FUNCTION_BLOCK "RD_PR_GantryUnload_Seqv25"   // FB2, LAD
VERSION : 0.1
// stored: AutoNumber true, IsIECCheckEnabled false, UDAEnableTagReadback false
   VAR_INPUT
      iAutoRunning : Bool;
      iCenteringSlideAtHome : Bool;
      iCenteringSlideAtWork : Bool;
      iDistSenHighLimit : Int;
      iDistSenLowLimit : Int;
      iDistSensorIP : Int;
      iDryCycleWithoutPal : Bool;
      iGantryOutofZone : Bool;
      iGantryPickOver : Bool;
      iPCAckZero : Bool;
      iPCBypass : Bool;
      iPCDataReadOver : Bool;
      iPCDataWriteOver : Bool;
      iPalletPresent : Bool;
      iProcessStart : Bool;
      iReset_fault : Bool;
      iRetryPB : Bool;
      iScanErr : Bool;
      iScanOver : Bool;
      iScannerBypass : Bool;
      iSstMode : Bool;
      iSstPB : Bool;
   END_VAR
   VAR_OUTPUT
      qCenteringSlideAdvance : Bool;
      qCenteringSlideRetract : Bool;
      qCheckDistance : Bool;
      qGantryOkToUnload : Bool;
      qMsg : Array[0..2] of Bool;
      qPCReadCmd : Bool;
      qPCUploadCmd : Bool;
      qProcessOver : Bool;
      qScanCmd : Bool;
   END_VAR
   VAR DB_SPECIFIC
      StateNo : Int;
      s44_WaitResetRelease : Bool;
      s44_WaitResetRelease_T1 : Bool;
      s45_WaitGantryOutZone : Bool;
      s45_WaitGantryOutZone_T1 : Bool;
      s46_ChkStationHome : Bool;
      s46_ChkStationHome_T1 : Bool;
      s46_ChkStationHome_T2 : Bool;
      s47_WaitProcStartPZR : Bool;
      s47_WaitProcStartPZR_T1 : Bool;
      s48_ChkRecovery : Bool;
      s48_ChkRecovery_T1 : Bool;
      s48_ChkRecovery_T2 : Bool;
      s48_ChkRecovery_T3 : Bool;
      s49_WaitCentSlideAdv : Bool;
      s49_WaitCentSlideAdv_T1 : Bool;
      s50_WaitDistSensorFB : Bool;
      s50_WaitDistSensorFB_T1 : Bool;
      s51_WaitCentSlideRet : Bool;
      s51_WaitCentSlideRet_T1 : Bool;
      s52_WaitScanOver : Bool;
      s52_WaitScanOver_T1 : Bool;
      s52_WaitScanOver_T2 : Bool;
      s53_ChkDistOkWithPC : Bool;
      s53_ChkDistOkWithPC_T1 : Bool;
      s53_ChkDistOkWithPC_T2 : Bool;
      s54_WaitGantryUnload : Bool;
      s54_WaitGantryUnload_T1 : Bool;
      s55_WaitGantryUnldOvr : Bool;
      s55_WaitGantryUnldOvr_T1 : Bool;
      s56_WaitGantryOutZone : Bool;
      s56_WaitGantryOutZone_T1 : Bool;
      s57_ChkReelAbsentConv : Bool;
      s57_ChkReelAbsentConv_T1 : Bool;
      s58_WaitProcStartLow : Bool;
      s58_WaitProcStartLow_T1 : Bool;
      s61_ChkMeasDiamTol : Bool;
      s61_ChkMeasDiamTol_T1 : Bool;
      s61_ChkMeasDiamTol_T2 : Bool;
      s62_WaitPCAckZero : Bool;
      s62_WaitPCAckZero_T1 : Bool;
      s63_WaitDataWritePC : Bool;
      s63_WaitDataWritePC_T1 : Bool;
      s64_WaitOperatorIntv : Bool;
      s64_WaitOperatorIntv_T1 : Bool;
      s65_ChkScanRetryOver : Bool;
      s65_ChkScanRetryOver_T1 : Bool;
      s65_ChkScanRetryOver_T2 : Bool;
      s66_WaitOperatorDecis : Bool;
      s66_WaitOperatorDecis_T1 : Bool;
      s67_WaitCentSlideRet : Bool;
      s67_WaitCentSlideRet_T1 : Bool;
      s68_WaitPCAckZeroRead : Bool;
      s68_WaitPCAckZeroRead_T1 : Bool;
      s69_WaitDataReadPC : Bool;
      s69_WaitDataReadPC_T1 : Bool;
      sDistanceHighLimit : Int;
      sDistanceLowLimit : Int;
      sRecoveryInt : Int;
      sScanRetryCount : Int;
      sSst : Bool;
      sSstPulse : Bool;
      sSstRise : Bool;
   END_VAR
   VAR_TEMP
      tOne : Bool;
   END_VAR
   VAR_TEMP   // added for the SCL form of the ladder/FBD networks
      _w1 : Bool;
   END_VAR
BEGIN

REGION Network 1
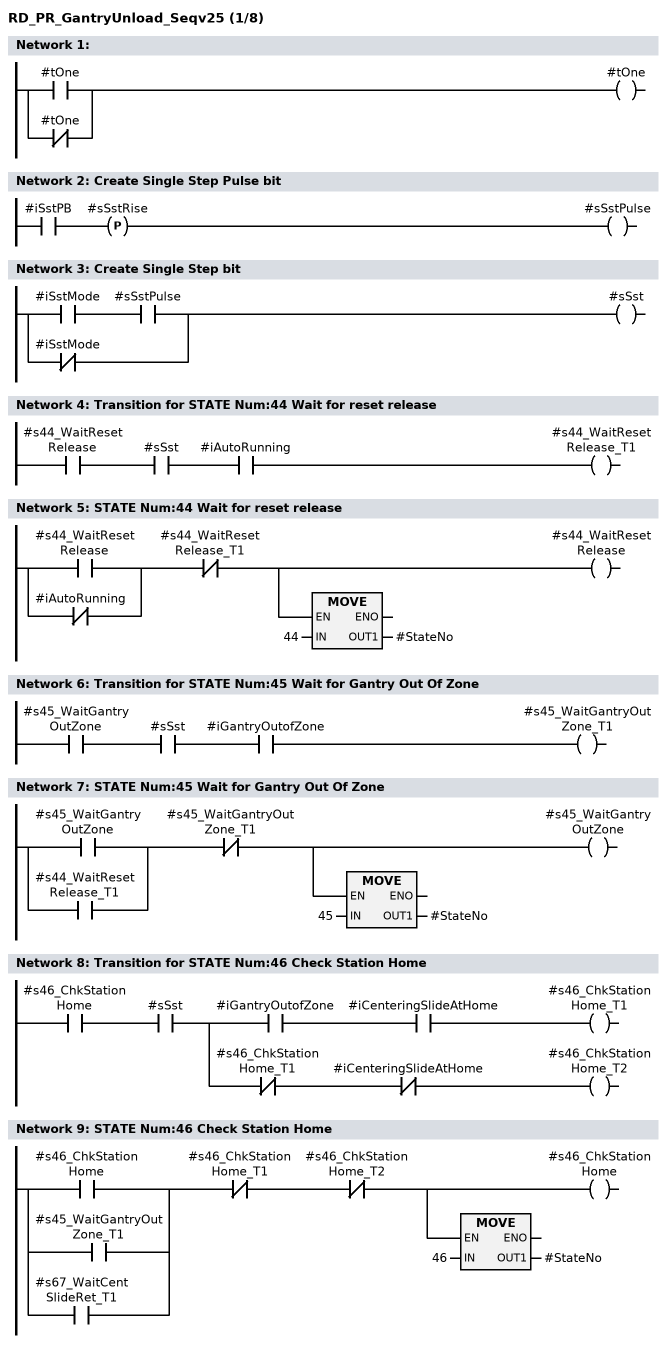
   RUNG wire#powerrail
      Contact( #tOne )
      wire#w1
      Coil( #tOne )
   END_RUNG
   RUNG wire#powerrail
      I_Contact( #tOne )
   END_RUNG wire#w1
   // the same network as SCL:
   #tOne := #tOne OR NOT #tOne;
END_REGION

REGION Network 2: Create Single Step Pulse bit
   RUNG wire#powerrail
      Contact( #iSstPB )
      P_Trig( #sSstRise )
      Coil( #sSstPulse )
   END_RUNG
   // the same network as SCL:
   #_w1 := #iSstPB AND NOT #sSstRise;   // rising edge
   #sSstRise := #iSstPB;
   #sSstPulse := #_w1;
END_REGION

REGION Network 3: Create Single Step bit
   RUNG wire#powerrail
      Contact( #iSstMode )
      Contact( #sSstPulse )
      wire#w1
      Coil( #sSst )
   END_RUNG
   RUNG wire#powerrail
      I_Contact( #iSstMode )
   END_RUNG wire#w1
   // the same network as SCL:
   #sSst := (#iSstMode AND #sSstPulse) OR NOT #iSstMode;
END_REGION

REGION Network 4: Transition for STATE Num:44 Wait for reset release
   RUNG wire#powerrail
      Contact( #s44_WaitResetRelease )
      Contact( #sSst )
      Contact( #iAutoRunning )
      Coil( #s44_WaitResetRelease_T1 )
   END_RUNG
   // the same network as SCL:
   #s44_WaitResetRelease_T1 := #s44_WaitResetRelease AND #sSst AND #iAutoRunning;
END_REGION

REGION Network 5: STATE Num:44 Wait for reset release
   RUNG wire#powerrail
      Contact( #s44_WaitResetRelease )
      wire#w1
      I_Contact( #s44_WaitResetRelease_T1 )
      wire#w2
      Coil( #s44_WaitResetRelease )
   END_RUNG
   RUNG wire#powerrail
      I_Contact( #iAutoRunning )
   END_RUNG wire#w1
   RUNG wire#w2
      { S7_GenerateENO := "TRUE" } Move(in := 44, out1 => #StateNo)
   END_RUNG
   // the same network as SCL:
   #s44_WaitResetRelease := (#s44_WaitResetRelease OR NOT #iAutoRunning) AND NOT #s44_WaitResetRelease_T1;
   IF #s44_WaitResetRelease THEN #StateNo := 44; END_IF;
END_REGION

REGION Network 6: Transition for STATE Num:45 Wait for Gantry Out Of Zone
   RUNG wire#powerrail
      Contact( #s45_WaitGantryOutZone )
      Contact( #sSst )
      Contact( #iGantryOutofZone )
      Coil( #s45_WaitGantryOutZone_T1 )
   END_RUNG
   // the same network as SCL:
   #s45_WaitGantryOutZone_T1 := #s45_WaitGantryOutZone AND #sSst AND #iGantryOutofZone;
END_REGION

REGION Network 7: STATE Num:45 Wait for Gantry Out Of Zone
   RUNG wire#powerrail
      Contact( #s45_WaitGantryOutZone )
      wire#w1
      I_Contact( #s45_WaitGantryOutZone_T1 )
      wire#w2
      Coil( #s45_WaitGantryOutZone )
   END_RUNG
   RUNG wire#powerrail
      Contact( #s44_WaitResetRelease_T1 )
   END_RUNG wire#w1
   RUNG wire#w2
      { S7_GenerateENO := "TRUE" } Move(in := 45, out1 => #StateNo)
   END_RUNG
   // the same network as SCL:
   #s45_WaitGantryOutZone := (#s45_WaitGantryOutZone OR #s44_WaitResetRelease_T1) AND NOT #s45_WaitGantryOutZone_T1;
   IF #s45_WaitGantryOutZone THEN #StateNo := 45; END_IF;
END_REGION

REGION Network 8: Transition for STATE Num:46 Check Station Home
   RUNG wire#powerrail
      Contact( #s46_ChkStationHome )
      Contact( #sSst )
      wire#w1
      Contact( #iGantryOutofZone )
      Contact( #iCenteringSlideAtHome )
      Coil( #s46_ChkStationHome_T1 )
   END_RUNG
   RUNG wire#w1
      I_Contact( #s46_ChkStationHome_T1 )
      I_Contact( #iCenteringSlideAtHome )
      Coil( #s46_ChkStationHome_T2 )
   END_RUNG
   // the same network as SCL:
   #_w1 := #s46_ChkStationHome AND #sSst;
   #s46_ChkStationHome_T1 := #_w1 AND #iGantryOutofZone AND #iCenteringSlideAtHome;
   #s46_ChkStationHome_T2 := #_w1 AND NOT #s46_ChkStationHome_T1 AND NOT #iCenteringSlideAtHome;
END_REGION

REGION Network 9: STATE Num:46 Check Station Home
   RUNG wire#powerrail
      Contact( #s46_ChkStationHome )
      wire#w1
      I_Contact( #s46_ChkStationHome_T1 )
      I_Contact( #s46_ChkStationHome_T2 )
      wire#w2
      Coil( #s46_ChkStationHome )
   END_RUNG
   RUNG wire#powerrail
      Contact( #s45_WaitGantryOutZone_T1 )
   END_RUNG wire#w1
   RUNG wire#powerrail
      Contact( #s67_WaitCentSlideRet_T1 )
   END_RUNG wire#w1
   RUNG wire#w2
      { S7_GenerateENO := "TRUE" } Move(in := 46, out1 => #StateNo)
   END_RUNG
   // the same network as SCL:
   #s46_ChkStationHome := (#s46_ChkStationHome OR #s45_WaitGantryOutZone_T1 OR #s67_WaitCentSlideRet_T1) AND NOT #s46_ChkStationHome_T1 AND NOT #s46_ChkStationHome_T2;
   IF #s46_ChkStationHome THEN #StateNo := 46; END_IF;
END_REGION

REGION Network 10: Transition for STATE Num:47 Wait for Process Start From PZR
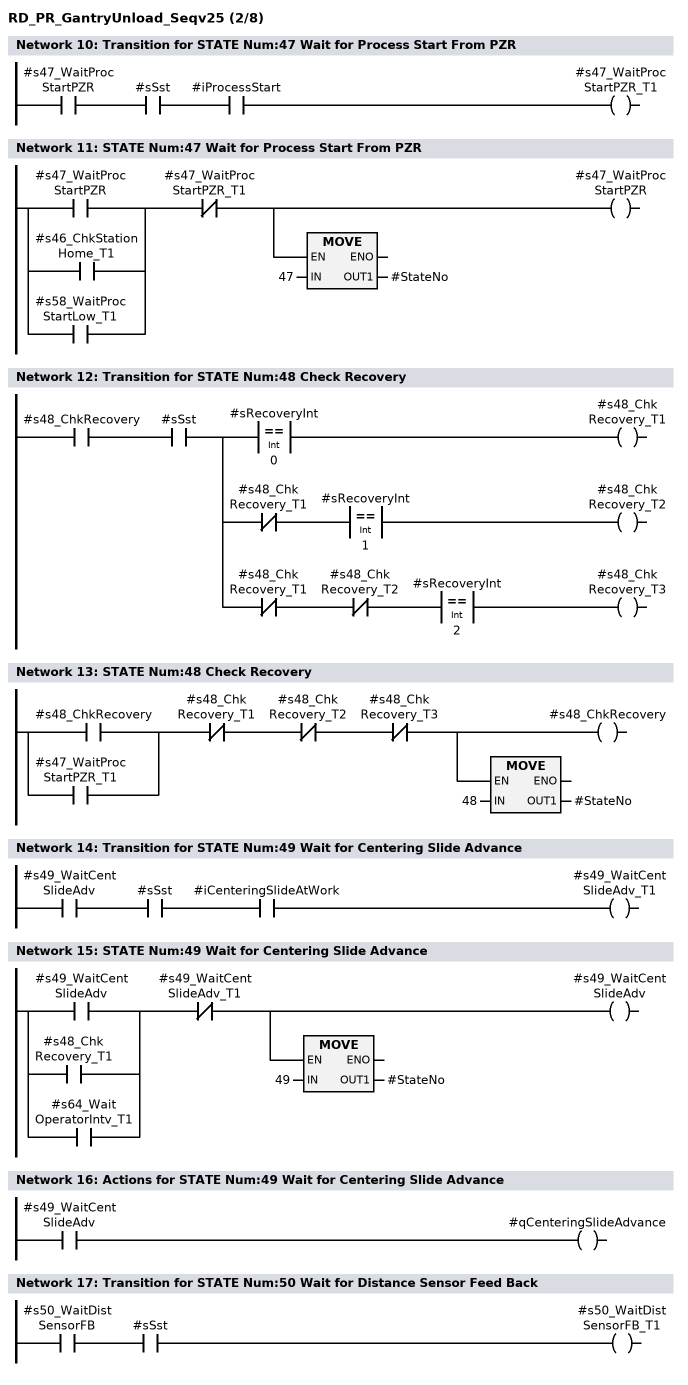
   RUNG wire#powerrail
      Contact( #s47_WaitProcStartPZR )
      Contact( #sSst )
      Contact( #iProcessStart )
      Coil( #s47_WaitProcStartPZR_T1 )
   END_RUNG
   // the same network as SCL:
   #s47_WaitProcStartPZR_T1 := #s47_WaitProcStartPZR AND #sSst AND #iProcessStart;
END_REGION

REGION Network 11: STATE Num:47 Wait for Process Start From PZR
   RUNG wire#powerrail
      Contact( #s47_WaitProcStartPZR )
      wire#w1
      I_Contact( #s47_WaitProcStartPZR_T1 )
      wire#w2
      Coil( #s47_WaitProcStartPZR )
   END_RUNG
   RUNG wire#powerrail
      Contact( #s46_ChkStationHome_T1 )
   END_RUNG wire#w1
   RUNG wire#powerrail
      Contact( #s58_WaitProcStartLow_T1 )
   END_RUNG wire#w1
   RUNG wire#w2
      { S7_GenerateENO := "TRUE" } Move(in := 47, out1 => #StateNo)
   END_RUNG
   // the same network as SCL:
   #s47_WaitProcStartPZR := (#s47_WaitProcStartPZR OR #s46_ChkStationHome_T1 OR #s58_WaitProcStartLow_T1) AND NOT #s47_WaitProcStartPZR_T1;
   IF #s47_WaitProcStartPZR THEN #StateNo := 47; END_IF;
END_REGION

REGION Network 12: Transition for STATE Num:48 Check Recovery
   RUNG wire#powerrail
      Contact( #s48_ChkRecovery )
      Contact( #sSst )
      wire#w1
      { S7_Templates := "SrcType := Int" } EQ_Contact(in1 := #sRecoveryInt, in2 := 0)
      Coil( #s48_ChkRecovery_T1 )
   END_RUNG
   RUNG wire#w1
      I_Contact( #s48_ChkRecovery_T1 )
      { S7_Templates := "SrcType := Int" } EQ_Contact(in1 := #sRecoveryInt, in2 := 1)
      Coil( #s48_ChkRecovery_T2 )
   END_RUNG
   RUNG wire#w1
      I_Contact( #s48_ChkRecovery_T1 )
      I_Contact( #s48_ChkRecovery_T2 )
      { S7_Templates := "SrcType := Int" } EQ_Contact(in1 := #sRecoveryInt, in2 := 2)
      Coil( #s48_ChkRecovery_T3 )
   END_RUNG
   // the same network as SCL:
   #_w1 := #s48_ChkRecovery AND #sSst;
   #s48_ChkRecovery_T1 := #_w1 AND (#sRecoveryInt = 0);
   #s48_ChkRecovery_T2 := #_w1 AND NOT #s48_ChkRecovery_T1 AND (#sRecoveryInt = 1);
   #s48_ChkRecovery_T3 := #_w1 AND NOT #s48_ChkRecovery_T1 AND NOT #s48_ChkRecovery_T2 AND (#sRecoveryInt = 2);
END_REGION

REGION Network 13: STATE Num:48 Check Recovery
   RUNG wire#powerrail
      Contact( #s48_ChkRecovery )
      wire#w1
      I_Contact( #s48_ChkRecovery_T1 )
      I_Contact( #s48_ChkRecovery_T2 )
      I_Contact( #s48_ChkRecovery_T3 )
      wire#w2
      Coil( #s48_ChkRecovery )
   END_RUNG
   RUNG wire#powerrail
      Contact( #s47_WaitProcStartPZR_T1 )
   END_RUNG wire#w1
   RUNG wire#w2
      { S7_GenerateENO := "TRUE" } Move(in := 48, out1 => #StateNo)
   END_RUNG
   // the same network as SCL:
   #s48_ChkRecovery := (#s48_ChkRecovery OR #s47_WaitProcStartPZR_T1) AND NOT #s48_ChkRecovery_T1 AND NOT #s48_ChkRecovery_T2 AND NOT #s48_ChkRecovery_T3;
   IF #s48_ChkRecovery THEN #StateNo := 48; END_IF;
END_REGION

REGION Network 14: Transition for STATE Num:49 Wait for Centering Slide Advance
   RUNG wire#powerrail
      Contact( #s49_WaitCentSlideAdv )
      Contact( #sSst )
      Contact( #iCenteringSlideAtWork )
      Coil( #s49_WaitCentSlideAdv_T1 )
   END_RUNG
   // the same network as SCL:
   #s49_WaitCentSlideAdv_T1 := #s49_WaitCentSlideAdv AND #sSst AND #iCenteringSlideAtWork;
END_REGION

REGION Network 15: STATE Num:49 Wait for Centering Slide Advance
   RUNG wire#powerrail
      Contact( #s49_WaitCentSlideAdv )
      wire#w1
      I_Contact( #s49_WaitCentSlideAdv_T1 )
      wire#w2
      Coil( #s49_WaitCentSlideAdv )
   END_RUNG
   RUNG wire#powerrail
      Contact( #s48_ChkRecovery_T1 )
   END_RUNG wire#w1
   RUNG wire#powerrail
      Contact( #s64_WaitOperatorIntv_T1 )
   END_RUNG wire#w1
   RUNG wire#w2
      { S7_GenerateENO := "TRUE" } Move(in := 49, out1 => #StateNo)
   END_RUNG
   // the same network as SCL:
   #s49_WaitCentSlideAdv := (#s49_WaitCentSlideAdv OR #s48_ChkRecovery_T1 OR #s64_WaitOperatorIntv_T1) AND NOT #s49_WaitCentSlideAdv_T1;
   IF #s49_WaitCentSlideAdv THEN #StateNo := 49; END_IF;
END_REGION

REGION Network 16: Actions for STATE Num:49 Wait for Centering Slide Advance
   RUNG wire#powerrail
      Contact( #s49_WaitCentSlideAdv )
      Coil( #qCenteringSlideAdvance )
   END_RUNG
   // the same network as SCL:
   #qCenteringSlideAdvance := #s49_WaitCentSlideAdv;
END_REGION

REGION Network 17: Transition for STATE Num:50 Wait for Distance Sensor Feed Back
   RUNG wire#powerrail
      Contact( #s50_WaitDistSensorFB )
      Contact( #sSst )
      Coil( #s50_WaitDistSensorFB_T1 )
   END_RUNG
   // the same network as SCL:
   #s50_WaitDistSensorFB_T1 := #s50_WaitDistSensorFB AND #sSst;
END_REGION

REGION Network 18: STATE Num:50 Wait for Distance Sensor Feed Back
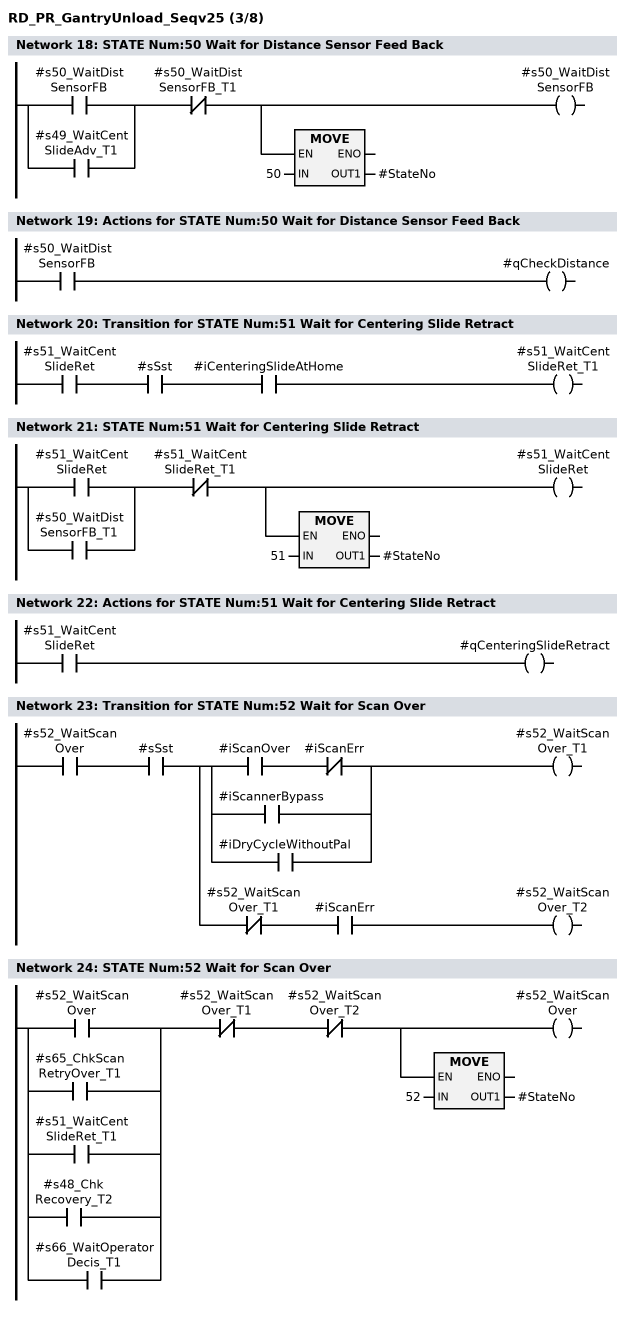
   RUNG wire#powerrail
      Contact( #s50_WaitDistSensorFB )
      wire#w1
      I_Contact( #s50_WaitDistSensorFB_T1 )
      wire#w2
      Coil( #s50_WaitDistSensorFB )
   END_RUNG
   RUNG wire#powerrail
      Contact( #s49_WaitCentSlideAdv_T1 )
   END_RUNG wire#w1
   RUNG wire#w2
      { S7_GenerateENO := "TRUE" } Move(in := 50, out1 => #StateNo)
   END_RUNG
   // the same network as SCL:
   #s50_WaitDistSensorFB := (#s50_WaitDistSensorFB OR #s49_WaitCentSlideAdv_T1) AND NOT #s50_WaitDistSensorFB_T1;
   IF #s50_WaitDistSensorFB THEN #StateNo := 50; END_IF;
END_REGION

REGION Network 19: Actions for STATE Num:50 Wait for Distance Sensor Feed Back
   RUNG wire#powerrail
      Contact( #s50_WaitDistSensorFB )
      Coil( #qCheckDistance )
   END_RUNG
   // the same network as SCL:
   #qCheckDistance := #s50_WaitDistSensorFB;
END_REGION

REGION Network 20: Transition for STATE Num:51 Wait for Centering Slide Retract
   RUNG wire#powerrail
      Contact( #s51_WaitCentSlideRet )
      Contact( #sSst )
      Contact( #iCenteringSlideAtHome )
      Coil( #s51_WaitCentSlideRet_T1 )
   END_RUNG
   // the same network as SCL:
   #s51_WaitCentSlideRet_T1 := #s51_WaitCentSlideRet AND #sSst AND #iCenteringSlideAtHome;
END_REGION

REGION Network 21: STATE Num:51 Wait for Centering Slide Retract
   RUNG wire#powerrail
      Contact( #s51_WaitCentSlideRet )
      wire#w1
      I_Contact( #s51_WaitCentSlideRet_T1 )
      wire#w2
      Coil( #s51_WaitCentSlideRet )
   END_RUNG
   RUNG wire#powerrail
      Contact( #s50_WaitDistSensorFB_T1 )
   END_RUNG wire#w1
   RUNG wire#w2
      { S7_GenerateENO := "TRUE" } Move(in := 51, out1 => #StateNo)
   END_RUNG
   // the same network as SCL:
   #s51_WaitCentSlideRet := (#s51_WaitCentSlideRet OR #s50_WaitDistSensorFB_T1) AND NOT #s51_WaitCentSlideRet_T1;
   IF #s51_WaitCentSlideRet THEN #StateNo := 51; END_IF;
END_REGION

REGION Network 22: Actions for STATE Num:51 Wait for Centering Slide Retract
   RUNG wire#powerrail
      Contact( #s51_WaitCentSlideRet )
      Coil( #qCenteringSlideRetract )
   END_RUNG
   // the same network as SCL:
   #qCenteringSlideRetract := #s51_WaitCentSlideRet;
END_REGION

REGION Network 23: Transition for STATE Num:52 Wait for Scan Over
   RUNG wire#powerrail
      Contact( #s52_WaitScanOver )
      Contact( #sSst )
      wire#w1
      Contact( #iScanOver )
      I_Contact( #iScanErr )
      wire#w2
      Coil( #s52_WaitScanOver_T1 )
   END_RUNG
   RUNG wire#w1
      Contact( #iScannerBypass )
   END_RUNG wire#w2
   RUNG wire#w1
      Contact( #iDryCycleWithoutPal )
   END_RUNG wire#w2
   RUNG wire#w1
      I_Contact( #s52_WaitScanOver_T1 )
      Contact( #iScanErr )
      Coil( #s52_WaitScanOver_T2 )
   END_RUNG
   // the same network as SCL:
   #_w1 := #s52_WaitScanOver AND #sSst;
   #s52_WaitScanOver_T1 := #_w1 AND ((#iScanOver AND NOT #iScanErr) OR #iScannerBypass OR #iDryCycleWithoutPal);
   #s52_WaitScanOver_T2 := #_w1 AND NOT #s52_WaitScanOver_T1 AND #iScanErr;
END_REGION

REGION Network 24: STATE Num:52 Wait for Scan Over
   RUNG wire#powerrail
      Contact( #s52_WaitScanOver )
      wire#w1
      I_Contact( #s52_WaitScanOver_T1 )
      I_Contact( #s52_WaitScanOver_T2 )
      wire#w2
      Coil( #s52_WaitScanOver )
   END_RUNG
   RUNG wire#powerrail
      Contact( #s65_ChkScanRetryOver_T1 )
   END_RUNG wire#w1
   RUNG wire#powerrail
      Contact( #s51_WaitCentSlideRet_T1 )
   END_RUNG wire#w1
   RUNG wire#powerrail
      Contact( #s48_ChkRecovery_T2 )
   END_RUNG wire#w1
   RUNG wire#powerrail
      Contact( #s66_WaitOperatorDecis_T1 )
   END_RUNG wire#w1
   RUNG wire#w2
      { S7_GenerateENO := "TRUE" } Move(in := 52, out1 => #StateNo)
   END_RUNG
   // the same network as SCL:
   #s52_WaitScanOver := (#s52_WaitScanOver OR #s65_ChkScanRetryOver_T1 OR #s51_WaitCentSlideRet_T1 OR #s48_ChkRecovery_T2 OR #s66_WaitOperatorDecis_T1) AND NOT #s52_WaitScanOver_T1 AND NOT #s52_WaitScanOver_T2;
   IF #s52_WaitScanOver THEN #StateNo := 52; END_IF;
END_REGION

REGION Network 25: Actions for STATE Num:52 Wait for Scan Over
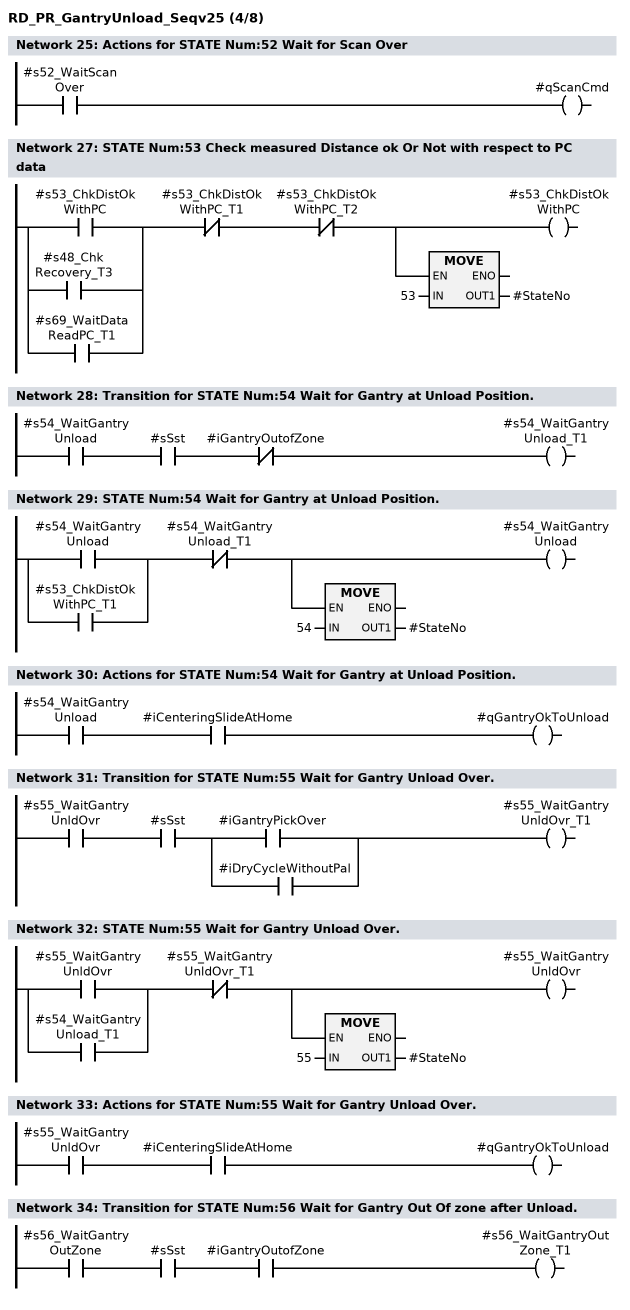
   RUNG wire#powerrail
      Contact( #s52_WaitScanOver )
      Coil( #qScanCmd )
   END_RUNG
   // the same network as SCL:
   #qScanCmd := #s52_WaitScanOver;
END_REGION

NETWORK
TITLE = Transition for STATE Num:53 Check measured Distance ok Or Not with respect to PC data
      A     #s53_ChkDistOkWithPC;
      A     #sSst;
      =     %L1.0;
      A     %L1.0;
      A(;
      L     #iDistSensorIP;
      L     #sDistanceLowLimit;
      >=R;
      );
      O(;
      L     #iDistSensorIP;
      L     #sDistanceHighLimit;
      <=R;
      );
      =     #s53_ChkDistOkWithPC_T1;
      A     %L1.0;
      AN    #s53_ChkDistOkWithPC_T1;
      A(;
      L     #iDistSensorIP;
      L     #sDistanceLowLimit;
      <R;
      );
      O(;
      L     #iDistSensorIP;
      L     #sDistanceHighLimit;
      >R;
      );
      =     #s53_ChkDistOkWithPC_T2;

REGION Network 27: STATE Num:53 Check measured Distance ok Or Not with respect to PC data
   RUNG wire#powerrail
      Contact( #s53_ChkDistOkWithPC )
      wire#w1
      I_Contact( #s53_ChkDistOkWithPC_T1 )
      I_Contact( #s53_ChkDistOkWithPC_T2 )
      wire#w2
      Coil( #s53_ChkDistOkWithPC )
   END_RUNG
   RUNG wire#powerrail
      Contact( #s48_ChkRecovery_T3 )
   END_RUNG wire#w1
   RUNG wire#powerrail
      Contact( #s69_WaitDataReadPC_T1 )
   END_RUNG wire#w1
   RUNG wire#w2
      { S7_GenerateENO := "TRUE" } Move(in := 53, out1 => #StateNo)
   END_RUNG
   // the same network as SCL:
   #s53_ChkDistOkWithPC := (#s53_ChkDistOkWithPC OR #s48_ChkRecovery_T3 OR #s69_WaitDataReadPC_T1) AND NOT #s53_ChkDistOkWithPC_T1 AND NOT #s53_ChkDistOkWithPC_T2;
   IF #s53_ChkDistOkWithPC THEN #StateNo := 53; END_IF;
END_REGION

REGION Network 28: Transition for STATE Num:54 Wait for Gantry at Unload Position.
   RUNG wire#powerrail
      Contact( #s54_WaitGantryUnload )
      Contact( #sSst )
      I_Contact( #iGantryOutofZone )
      Coil( #s54_WaitGantryUnload_T1 )
   END_RUNG
   // the same network as SCL:
   #s54_WaitGantryUnload_T1 := #s54_WaitGantryUnload AND #sSst AND NOT #iGantryOutofZone;
END_REGION

REGION Network 29: STATE Num:54 Wait for Gantry at Unload Position.
   RUNG wire#powerrail
      Contact( #s54_WaitGantryUnload )
      wire#w1
      I_Contact( #s54_WaitGantryUnload_T1 )
      wire#w2
      Coil( #s54_WaitGantryUnload )
   END_RUNG
   RUNG wire#powerrail
      Contact( #s53_ChkDistOkWithPC_T1 )
   END_RUNG wire#w1
   RUNG wire#w2
      { S7_GenerateENO := "TRUE" } Move(in := 54, out1 => #StateNo)
   END_RUNG
   // the same network as SCL:
   #s54_WaitGantryUnload := (#s54_WaitGantryUnload OR #s53_ChkDistOkWithPC_T1) AND NOT #s54_WaitGantryUnload_T1;
   IF #s54_WaitGantryUnload THEN #StateNo := 54; END_IF;
END_REGION

REGION Network 30: Actions for STATE Num:54 Wait for Gantry at Unload Position.
   RUNG wire#powerrail
      Contact( #s54_WaitGantryUnload )
      Contact( #iCenteringSlideAtHome )
      Coil( #qGantryOkToUnload )
   END_RUNG
   // the same network as SCL:
   #qGantryOkToUnload := #s54_WaitGantryUnload AND #iCenteringSlideAtHome;
END_REGION

REGION Network 31: Transition for STATE Num:55 Wait for Gantry Unload Over.
   RUNG wire#powerrail
      Contact( #s55_WaitGantryUnldOvr )
      Contact( #sSst )
      wire#w1
      Contact( #iGantryPickOver )
      wire#w2
      Coil( #s55_WaitGantryUnldOvr_T1 )
   END_RUNG
   RUNG wire#w1
      Contact( #iDryCycleWithoutPal )
   END_RUNG wire#w2
   // the same network as SCL:
   #s55_WaitGantryUnldOvr_T1 := #s55_WaitGantryUnldOvr AND #sSst AND (#iGantryPickOver OR #iDryCycleWithoutPal);
END_REGION

REGION Network 32: STATE Num:55 Wait for Gantry Unload Over.
   RUNG wire#powerrail
      Contact( #s55_WaitGantryUnldOvr )
      wire#w1
      I_Contact( #s55_WaitGantryUnldOvr_T1 )
      wire#w2
      Coil( #s55_WaitGantryUnldOvr )
   END_RUNG
   RUNG wire#powerrail
      Contact( #s54_WaitGantryUnload_T1 )
   END_RUNG wire#w1
   RUNG wire#w2
      { S7_GenerateENO := "TRUE" } Move(in := 55, out1 => #StateNo)
   END_RUNG
   // the same network as SCL:
   #s55_WaitGantryUnldOvr := (#s55_WaitGantryUnldOvr OR #s54_WaitGantryUnload_T1) AND NOT #s55_WaitGantryUnldOvr_T1;
   IF #s55_WaitGantryUnldOvr THEN #StateNo := 55; END_IF;
END_REGION

REGION Network 33: Actions for STATE Num:55 Wait for Gantry Unload Over.
   RUNG wire#powerrail
      Contact( #s55_WaitGantryUnldOvr )
      Contact( #iCenteringSlideAtHome )
      Coil( #qGantryOkToUnload )
   END_RUNG
   // the same network as SCL:
   #qGantryOkToUnload := #s55_WaitGantryUnldOvr AND #iCenteringSlideAtHome;
END_REGION

REGION Network 34: Transition for STATE Num:56 Wait for Gantry Out Of zone after Unload.
   RUNG wire#powerrail
      Contact( #s56_WaitGantryOutZone )
      Contact( #sSst )
      Contact( #iGantryOutofZone )
      Coil( #s56_WaitGantryOutZone_T1 )
   END_RUNG
   // the same network as SCL:
   #s56_WaitGantryOutZone_T1 := #s56_WaitGantryOutZone AND #sSst AND #iGantryOutofZone;
END_REGION

REGION Network 35: STATE Num:56 Wait for Gantry Out Of zone after Unload.
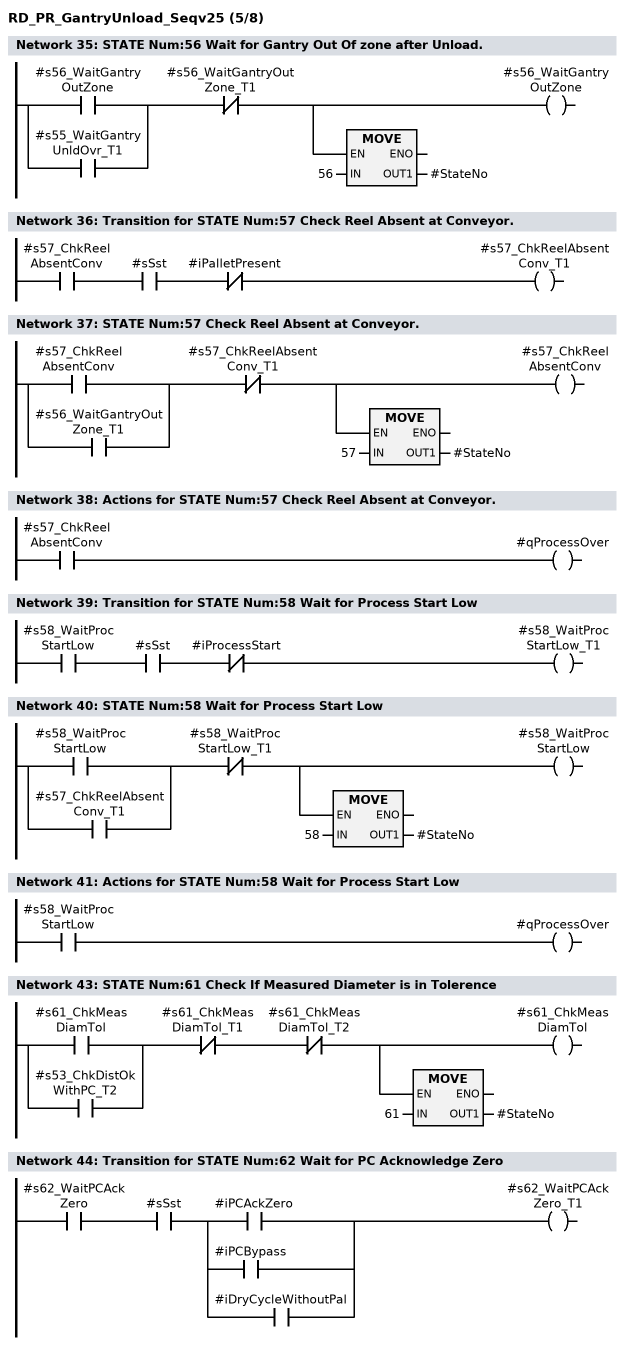
   RUNG wire#powerrail
      Contact( #s56_WaitGantryOutZone )
      wire#w1
      I_Contact( #s56_WaitGantryOutZone_T1 )
      wire#w2
      Coil( #s56_WaitGantryOutZone )
   END_RUNG
   RUNG wire#powerrail
      Contact( #s55_WaitGantryUnldOvr_T1 )
   END_RUNG wire#w1
   RUNG wire#w2
      { S7_GenerateENO := "TRUE" } Move(in := 56, out1 => #StateNo)
   END_RUNG
   // the same network as SCL:
   #s56_WaitGantryOutZone := (#s56_WaitGantryOutZone OR #s55_WaitGantryUnldOvr_T1) AND NOT #s56_WaitGantryOutZone_T1;
   IF #s56_WaitGantryOutZone THEN #StateNo := 56; END_IF;
END_REGION

REGION Network 36: Transition for STATE Num:57 Check Reel Absent at Conveyor.
   RUNG wire#powerrail
      Contact( #s57_ChkReelAbsentConv )
      Contact( #sSst )
      I_Contact( #iPalletPresent )
      Coil( #s57_ChkReelAbsentConv_T1 )
   END_RUNG
   // the same network as SCL:
   #s57_ChkReelAbsentConv_T1 := #s57_ChkReelAbsentConv AND #sSst AND NOT #iPalletPresent;
END_REGION

REGION Network 37: STATE Num:57 Check Reel Absent at Conveyor.
   RUNG wire#powerrail
      Contact( #s57_ChkReelAbsentConv )
      wire#w1
      I_Contact( #s57_ChkReelAbsentConv_T1 )
      wire#w2
      Coil( #s57_ChkReelAbsentConv )
   END_RUNG
   RUNG wire#powerrail
      Contact( #s56_WaitGantryOutZone_T1 )
   END_RUNG wire#w1
   RUNG wire#w2
      { S7_GenerateENO := "TRUE" } Move(in := 57, out1 => #StateNo)
   END_RUNG
   // the same network as SCL:
   #s57_ChkReelAbsentConv := (#s57_ChkReelAbsentConv OR #s56_WaitGantryOutZone_T1) AND NOT #s57_ChkReelAbsentConv_T1;
   IF #s57_ChkReelAbsentConv THEN #StateNo := 57; END_IF;
END_REGION

REGION Network 38: Actions for STATE Num:57 Check Reel Absent at Conveyor.
   RUNG wire#powerrail
      Contact( #s57_ChkReelAbsentConv )
      Coil( #qProcessOver )
   END_RUNG
   // the same network as SCL:
   #qProcessOver := #s57_ChkReelAbsentConv;
END_REGION

REGION Network 39: Transition for STATE Num:58 Wait for Process Start Low
   RUNG wire#powerrail
      Contact( #s58_WaitProcStartLow )
      Contact( #sSst )
      I_Contact( #iProcessStart )
      Coil( #s58_WaitProcStartLow_T1 )
   END_RUNG
   // the same network as SCL:
   #s58_WaitProcStartLow_T1 := #s58_WaitProcStartLow AND #sSst AND NOT #iProcessStart;
END_REGION

REGION Network 40: STATE Num:58 Wait for Process Start Low
   RUNG wire#powerrail
      Contact( #s58_WaitProcStartLow )
      wire#w1
      I_Contact( #s58_WaitProcStartLow_T1 )
      wire#w2
      Coil( #s58_WaitProcStartLow )
   END_RUNG
   RUNG wire#powerrail
      Contact( #s57_ChkReelAbsentConv_T1 )
   END_RUNG wire#w1
   RUNG wire#w2
      { S7_GenerateENO := "TRUE" } Move(in := 58, out1 => #StateNo)
   END_RUNG
   // the same network as SCL:
   #s58_WaitProcStartLow := (#s58_WaitProcStartLow OR #s57_ChkReelAbsentConv_T1) AND NOT #s58_WaitProcStartLow_T1;
   IF #s58_WaitProcStartLow THEN #StateNo := 58; END_IF;
END_REGION

REGION Network 41: Actions for STATE Num:58 Wait for Process Start Low
   RUNG wire#powerrail
      Contact( #s58_WaitProcStartLow )
      Coil( #qProcessOver )
   END_RUNG
   // the same network as SCL:
   #qProcessOver := #s58_WaitProcStartLow;
END_REGION

NETWORK
TITLE = Transition for STATE Num:61 Check If Measured Diameter is in Tolerence
      A     #s61_ChkMeasDiamTol;
      A     #sSst;
      =     %L1.0;
      A     %L1.0;
      A(;
      L     #iDistSenLowLimit;
      L     #iDistSensorIP;
      <=R;
      );
      O(;
      L     #iDistSensorIP;
      L     #iDistSenHighLimit;
      <=R;
      );
      =     #s61_ChkMeasDiamTol_T1;
      A     %L1.0;
      AN    #s61_ChkMeasDiamTol_T1;
      A(;
      L     #iDistSenLowLimit;
      L     #iDistSensorIP;
      >R;
      );
      O(;
      L     #iDistSensorIP;
      L     #iDistSenHighLimit;
      >R;
      );
      =     #s61_ChkMeasDiamTol_T2;

REGION Network 43: STATE Num:61 Check If Measured Diameter is in Tolerence
   RUNG wire#powerrail
      Contact( #s61_ChkMeasDiamTol )
      wire#w1
      I_Contact( #s61_ChkMeasDiamTol_T1 )
      I_Contact( #s61_ChkMeasDiamTol_T2 )
      wire#w2
      Coil( #s61_ChkMeasDiamTol )
   END_RUNG
   RUNG wire#powerrail
      Contact( #s53_ChkDistOkWithPC_T2 )
   END_RUNG wire#w1
   RUNG wire#w2
      { S7_GenerateENO := "TRUE" } Move(in := 61, out1 => #StateNo)
   END_RUNG
   // the same network as SCL:
   #s61_ChkMeasDiamTol := (#s61_ChkMeasDiamTol OR #s53_ChkDistOkWithPC_T2) AND NOT #s61_ChkMeasDiamTol_T1 AND NOT #s61_ChkMeasDiamTol_T2;
   IF #s61_ChkMeasDiamTol THEN #StateNo := 61; END_IF;
END_REGION

REGION Network 44: Transition for STATE Num:62 Wait for PC Acknowledge Zero
   RUNG wire#powerrail
      Contact( #s62_WaitPCAckZero )
      Contact( #sSst )
      wire#w1
      Contact( #iPCAckZero )
      wire#w2
      Coil( #s62_WaitPCAckZero_T1 )
   END_RUNG
   RUNG wire#w1
      Contact( #iPCBypass )
   END_RUNG wire#w2
   RUNG wire#w1
      Contact( #iDryCycleWithoutPal )
   END_RUNG wire#w2
   // the same network as SCL:
   #s62_WaitPCAckZero_T1 := #s62_WaitPCAckZero AND #sSst AND (#iPCAckZero OR #iPCBypass OR #iDryCycleWithoutPal);
END_REGION

REGION Network 45: STATE Num:62 Wait for PC Acknowledge Zero
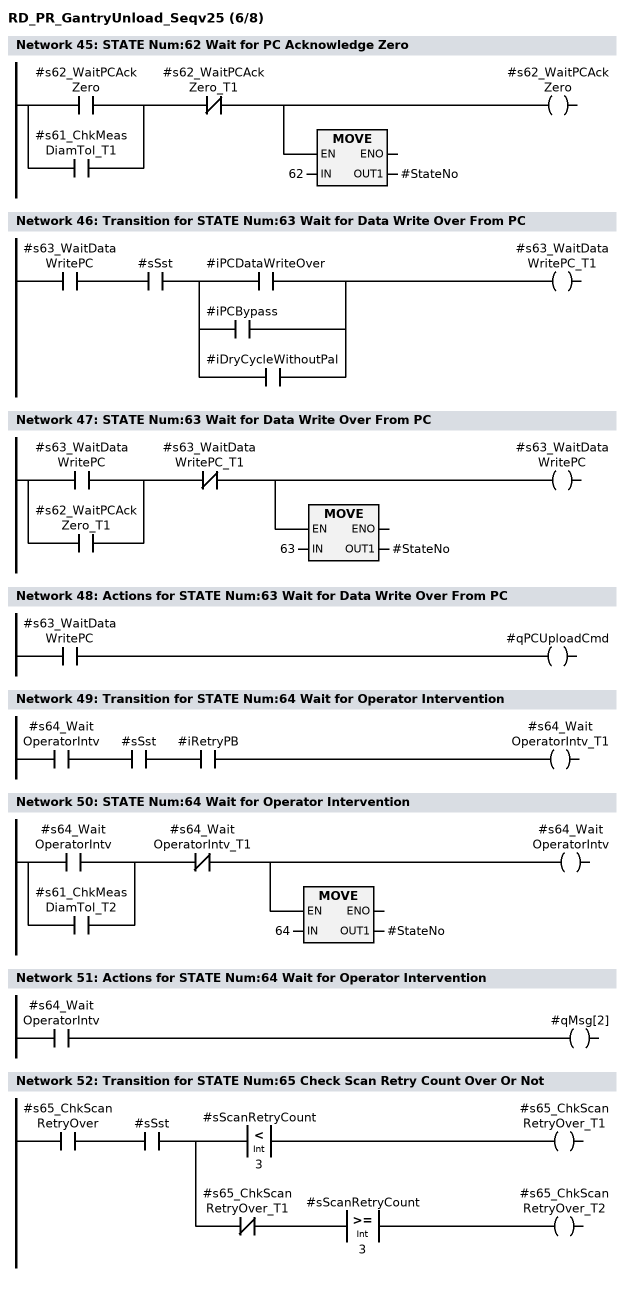
   RUNG wire#powerrail
      Contact( #s62_WaitPCAckZero )
      wire#w1
      I_Contact( #s62_WaitPCAckZero_T1 )
      wire#w2
      Coil( #s62_WaitPCAckZero )
   END_RUNG
   RUNG wire#powerrail
      Contact( #s61_ChkMeasDiamTol_T1 )
   END_RUNG wire#w1
   RUNG wire#w2
      { S7_GenerateENO := "TRUE" } Move(in := 62, out1 => #StateNo)
   END_RUNG
   // the same network as SCL:
   #s62_WaitPCAckZero := (#s62_WaitPCAckZero OR #s61_ChkMeasDiamTol_T1) AND NOT #s62_WaitPCAckZero_T1;
   IF #s62_WaitPCAckZero THEN #StateNo := 62; END_IF;
END_REGION

REGION Network 46: Transition for STATE Num:63 Wait for Data Write Over From PC
   RUNG wire#powerrail
      Contact( #s63_WaitDataWritePC )
      Contact( #sSst )
      wire#w1
      Contact( #iPCDataWriteOver )
      wire#w2
      Coil( #s63_WaitDataWritePC_T1 )
   END_RUNG
   RUNG wire#w1
      Contact( #iPCBypass )
   END_RUNG wire#w2
   RUNG wire#w1
      Contact( #iDryCycleWithoutPal )
   END_RUNG wire#w2
   // the same network as SCL:
   #s63_WaitDataWritePC_T1 := #s63_WaitDataWritePC AND #sSst AND (#iPCDataWriteOver OR #iPCBypass OR #iDryCycleWithoutPal);
END_REGION

REGION Network 47: STATE Num:63 Wait for Data Write Over From PC
   RUNG wire#powerrail
      Contact( #s63_WaitDataWritePC )
      wire#w1
      I_Contact( #s63_WaitDataWritePC_T1 )
      wire#w2
      Coil( #s63_WaitDataWritePC )
   END_RUNG
   RUNG wire#powerrail
      Contact( #s62_WaitPCAckZero_T1 )
   END_RUNG wire#w1
   RUNG wire#w2
      { S7_GenerateENO := "TRUE" } Move(in := 63, out1 => #StateNo)
   END_RUNG
   // the same network as SCL:
   #s63_WaitDataWritePC := (#s63_WaitDataWritePC OR #s62_WaitPCAckZero_T1) AND NOT #s63_WaitDataWritePC_T1;
   IF #s63_WaitDataWritePC THEN #StateNo := 63; END_IF;
END_REGION

REGION Network 48: Actions for STATE Num:63 Wait for Data Write Over From PC
   RUNG wire#powerrail
      Contact( #s63_WaitDataWritePC )
      Coil( #qPCUploadCmd )
   END_RUNG
   // the same network as SCL:
   #qPCUploadCmd := #s63_WaitDataWritePC;
END_REGION

REGION Network 49: Transition for STATE Num:64 Wait for Operator Intervention
   RUNG wire#powerrail
      Contact( #s64_WaitOperatorIntv )
      Contact( #sSst )
      Contact( #iRetryPB )
      Coil( #s64_WaitOperatorIntv_T1 )
   END_RUNG
   // the same network as SCL:
   #s64_WaitOperatorIntv_T1 := #s64_WaitOperatorIntv AND #sSst AND #iRetryPB;
END_REGION

REGION Network 50: STATE Num:64 Wait for Operator Intervention
   RUNG wire#powerrail
      Contact( #s64_WaitOperatorIntv )
      wire#w1
      I_Contact( #s64_WaitOperatorIntv_T1 )
      wire#w2
      Coil( #s64_WaitOperatorIntv )
   END_RUNG
   RUNG wire#powerrail
      Contact( #s61_ChkMeasDiamTol_T2 )
   END_RUNG wire#w1
   RUNG wire#w2
      { S7_GenerateENO := "TRUE" } Move(in := 64, out1 => #StateNo)
   END_RUNG
   // the same network as SCL:
   #s64_WaitOperatorIntv := (#s64_WaitOperatorIntv OR #s61_ChkMeasDiamTol_T2) AND NOT #s64_WaitOperatorIntv_T1;
   IF #s64_WaitOperatorIntv THEN #StateNo := 64; END_IF;
END_REGION

REGION Network 51: Actions for STATE Num:64 Wait for Operator Intervention
   RUNG wire#powerrail
      Contact( #s64_WaitOperatorIntv )
      Coil( #qMsg[2] )
   END_RUNG
   // the same network as SCL:
   #qMsg[2] := #s64_WaitOperatorIntv;
END_REGION

REGION Network 52: Transition for STATE Num:65 Check Scan Retry Count Over Or Not
   RUNG wire#powerrail
      Contact( #s65_ChkScanRetryOver )
      Contact( #sSst )
      wire#w1
      { S7_Templates := "SrcType := Int" } LT_Contact(in1 := #sScanRetryCount, in2 := 3)
      Coil( #s65_ChkScanRetryOver_T1 )
   END_RUNG
   RUNG wire#w1
      I_Contact( #s65_ChkScanRetryOver_T1 )
      { S7_Templates := "SrcType := Int" } GE_Contact(in1 := #sScanRetryCount, in2 := 3)
      Coil( #s65_ChkScanRetryOver_T2 )
   END_RUNG
   // the same network as SCL:
   #_w1 := #s65_ChkScanRetryOver AND #sSst;
   #s65_ChkScanRetryOver_T1 := #_w1 AND (#sScanRetryCount < 3);
   #s65_ChkScanRetryOver_T2 := #_w1 AND NOT #s65_ChkScanRetryOver_T1 AND (#sScanRetryCount >= 3);
END_REGION

REGION Network 53: STATE Num:65 Check Scan Retry Count Over Or Not
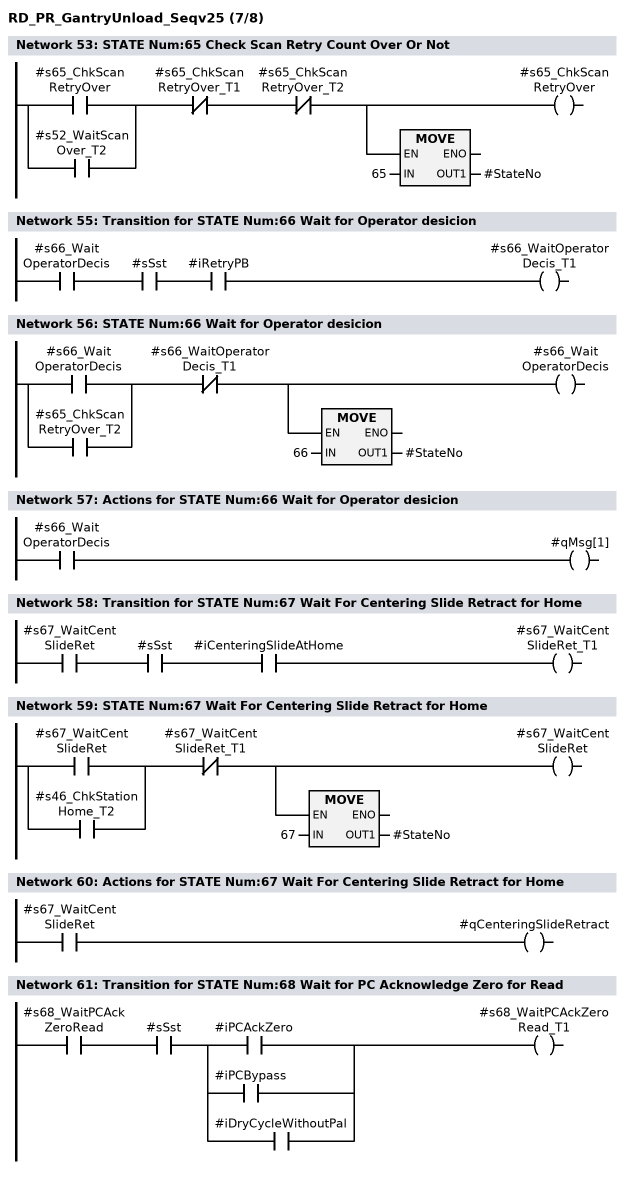
   RUNG wire#powerrail
      Contact( #s65_ChkScanRetryOver )
      wire#w1
      I_Contact( #s65_ChkScanRetryOver_T1 )
      I_Contact( #s65_ChkScanRetryOver_T2 )
      wire#w2
      Coil( #s65_ChkScanRetryOver )
   END_RUNG
   RUNG wire#powerrail
      Contact( #s52_WaitScanOver_T2 )
   END_RUNG wire#w1
   RUNG wire#w2
      { S7_GenerateENO := "TRUE" } Move(in := 65, out1 => #StateNo)
   END_RUNG
   // the same network as SCL:
   #s65_ChkScanRetryOver := (#s65_ChkScanRetryOver OR #s52_WaitScanOver_T2) AND NOT #s65_ChkScanRetryOver_T1 AND NOT #s65_ChkScanRetryOver_T2;
   IF #s65_ChkScanRetryOver THEN #StateNo := 65; END_IF;
END_REGION

NETWORK
TITLE = Actions for STATE Num:65 Check Scan Retry Count Over Or Not
      A     #s65_ChkScanRetryOver;
      A     #s65_ChkScanRetryOver_T1;
      L     #sScanRetryCount;
      L     1;
      +I;
      T     #sScanRetryCount;

REGION Network 55: Transition for STATE Num:66 Wait for Operator desicion
   RUNG wire#powerrail
      Contact( #s66_WaitOperatorDecis )
      Contact( #sSst )
      Contact( #iRetryPB )
      Coil( #s66_WaitOperatorDecis_T1 )
   END_RUNG
   // the same network as SCL:
   #s66_WaitOperatorDecis_T1 := #s66_WaitOperatorDecis AND #sSst AND #iRetryPB;
END_REGION

REGION Network 56: STATE Num:66 Wait for Operator desicion
   RUNG wire#powerrail
      Contact( #s66_WaitOperatorDecis )
      wire#w1
      I_Contact( #s66_WaitOperatorDecis_T1 )
      wire#w2
      Coil( #s66_WaitOperatorDecis )
   END_RUNG
   RUNG wire#powerrail
      Contact( #s65_ChkScanRetryOver_T2 )
   END_RUNG wire#w1
   RUNG wire#w2
      { S7_GenerateENO := "TRUE" } Move(in := 66, out1 => #StateNo)
   END_RUNG
   // the same network as SCL:
   #s66_WaitOperatorDecis := (#s66_WaitOperatorDecis OR #s65_ChkScanRetryOver_T2) AND NOT #s66_WaitOperatorDecis_T1;
   IF #s66_WaitOperatorDecis THEN #StateNo := 66; END_IF;
END_REGION

REGION Network 57: Actions for STATE Num:66 Wait for Operator desicion
   RUNG wire#powerrail
      Contact( #s66_WaitOperatorDecis )
      Coil( #qMsg[1] )
   END_RUNG
   // the same network as SCL:
   #qMsg[1] := #s66_WaitOperatorDecis;
END_REGION

REGION Network 58: Transition for STATE Num:67 Wait For Centering Slide Retract for Home
   RUNG wire#powerrail
      Contact( #s67_WaitCentSlideRet )
      Contact( #sSst )
      Contact( #iCenteringSlideAtHome )
      Coil( #s67_WaitCentSlideRet_T1 )
   END_RUNG
   // the same network as SCL:
   #s67_WaitCentSlideRet_T1 := #s67_WaitCentSlideRet AND #sSst AND #iCenteringSlideAtHome;
END_REGION

REGION Network 59: STATE Num:67 Wait For Centering Slide Retract for Home
   RUNG wire#powerrail
      Contact( #s67_WaitCentSlideRet )
      wire#w1
      I_Contact( #s67_WaitCentSlideRet_T1 )
      wire#w2
      Coil( #s67_WaitCentSlideRet )
   END_RUNG
   RUNG wire#powerrail
      Contact( #s46_ChkStationHome_T2 )
   END_RUNG wire#w1
   RUNG wire#w2
      { S7_GenerateENO := "TRUE" } Move(in := 67, out1 => #StateNo)
   END_RUNG
   // the same network as SCL:
   #s67_WaitCentSlideRet := (#s67_WaitCentSlideRet OR #s46_ChkStationHome_T2) AND NOT #s67_WaitCentSlideRet_T1;
   IF #s67_WaitCentSlideRet THEN #StateNo := 67; END_IF;
END_REGION

REGION Network 60: Actions for STATE Num:67 Wait For Centering Slide Retract for Home
   RUNG wire#powerrail
      Contact( #s67_WaitCentSlideRet )
      Coil( #qCenteringSlideRetract )
   END_RUNG
   // the same network as SCL:
   #qCenteringSlideRetract := #s67_WaitCentSlideRet;
END_REGION

REGION Network 61: Transition for STATE Num:68 Wait for PC Acknowledge Zero for Read
   RUNG wire#powerrail
      Contact( #s68_WaitPCAckZeroRead )
      Contact( #sSst )
      wire#w1
      Contact( #iPCAckZero )
      wire#w2
      Coil( #s68_WaitPCAckZeroRead_T1 )
   END_RUNG
   RUNG wire#w1
      Contact( #iPCBypass )
   END_RUNG wire#w2
   RUNG wire#w1
      Contact( #iDryCycleWithoutPal )
   END_RUNG wire#w2
   // the same network as SCL:
   #s68_WaitPCAckZeroRead_T1 := #s68_WaitPCAckZeroRead AND #sSst AND (#iPCAckZero OR #iPCBypass OR #iDryCycleWithoutPal);
END_REGION

REGION Network 62: STATE Num:68 Wait for PC Acknowledge Zero for Read
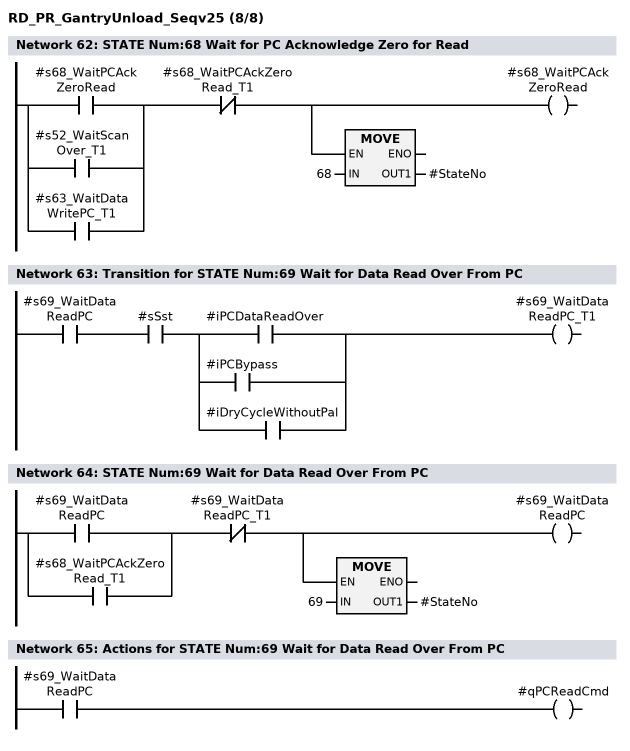
   RUNG wire#powerrail
      Contact( #s68_WaitPCAckZeroRead )
      wire#w1
      I_Contact( #s68_WaitPCAckZeroRead_T1 )
      wire#w2
      Coil( #s68_WaitPCAckZeroRead )
   END_RUNG
   RUNG wire#powerrail
      Contact( #s52_WaitScanOver_T1 )
   END_RUNG wire#w1
   RUNG wire#powerrail
      Contact( #s63_WaitDataWritePC_T1 )
   END_RUNG wire#w1
   RUNG wire#w2
      { S7_GenerateENO := "TRUE" } Move(in := 68, out1 => #StateNo)
   END_RUNG
   // the same network as SCL:
   #s68_WaitPCAckZeroRead := (#s68_WaitPCAckZeroRead OR #s52_WaitScanOver_T1 OR #s63_WaitDataWritePC_T1) AND NOT #s68_WaitPCAckZeroRead_T1;
   IF #s68_WaitPCAckZeroRead THEN #StateNo := 68; END_IF;
END_REGION

REGION Network 63: Transition for STATE Num:69 Wait for Data Read Over From PC
   RUNG wire#powerrail
      Contact( #s69_WaitDataReadPC )
      Contact( #sSst )
      wire#w1
      Contact( #iPCDataReadOver )
      wire#w2
      Coil( #s69_WaitDataReadPC_T1 )
   END_RUNG
   RUNG wire#w1
      Contact( #iPCBypass )
   END_RUNG wire#w2
   RUNG wire#w1
      Contact( #iDryCycleWithoutPal )
   END_RUNG wire#w2
   // the same network as SCL:
   #s69_WaitDataReadPC_T1 := #s69_WaitDataReadPC AND #sSst AND (#iPCDataReadOver OR #iPCBypass OR #iDryCycleWithoutPal);
END_REGION

REGION Network 64: STATE Num:69 Wait for Data Read Over From PC
   RUNG wire#powerrail
      Contact( #s69_WaitDataReadPC )
      wire#w1
      I_Contact( #s69_WaitDataReadPC_T1 )
      wire#w2
      Coil( #s69_WaitDataReadPC )
   END_RUNG
   RUNG wire#powerrail
      Contact( #s68_WaitPCAckZeroRead_T1 )
   END_RUNG wire#w1
   RUNG wire#w2
      { S7_GenerateENO := "TRUE" } Move(in := 69, out1 => #StateNo)
   END_RUNG
   // the same network as SCL:
   #s69_WaitDataReadPC := (#s69_WaitDataReadPC OR #s68_WaitPCAckZeroRead_T1) AND NOT #s69_WaitDataReadPC_T1;
   IF #s69_WaitDataReadPC THEN #StateNo := 69; END_IF;
END_REGION

REGION Network 65: Actions for STATE Num:69 Wait for Data Read Over From PC
   RUNG wire#powerrail
      Contact( #s69_WaitDataReadPC )
      Coil( #qPCReadCmd )
   END_RUNG
   // the same network as SCL:
   #qPCReadCmd := #s69_WaitDataReadPC;
END_REGION
END_FUNCTION_BLOCK

FUNCTION_BLOCK "S31808022001_Sequence_All_73b5c5_cfdfd9eb-ebd8-4267-a68e-df0ebcea3fa8 - Copy (2)_f93786"   // FB1, LAD
VERSION : 0.1
// stored: AutoNumber true, IsIECCheckEnabled false, UDAEnableTagReadback false
   VAR_INPUT
      iAutoRunning : Bool;
      iFaultReset : Bool;
      iOTS_Frm_Prev_TTDown : Bool;
      iOTS_Frm_Prev_TTUp : Bool;
      iPalletNtPrsntAtTTDown : Bool;
      iPalletNtPrsntAtTTUp : Bool;
      iPalletPrsnt_TTDown : Bool;
      iPalletPrsnt_TTUp : Bool;
      iPartReject : Bool;
      iRTR_Frm_Next_0DegTTUp : Bool;
      iRTR_Frm_Next_90DegTTUp : Bool;
      iRTR_Frm_Next_TTDown : Bool;
      iRecvAreaClr_TTDown : Bool;
      iRecvAreaClr_TTUp : Bool;
      iReset_fault : Bool;
      iRx_Frm_Prev_TTUp : Bool;
      iSstMode : Bool;
      iSstPB : Bool;
      iStprRaise_TTDown : Bool;
      iStprRaise_TTUp : Bool;
      iTTAt0Pos : Bool;
      iTTAt90Pos : Bool;
      iTTLocked : Bool;
      iTTUnlocked : Bool;
      iXferAreaClr_0DegTTDown : Bool;
      iXferAreaClr_0DegTTUp : Bool;
      iXferAreaClr_90DegTTUp : Bool;
   END_VAR
   VAR_OUTPUT
      qConvRun_TTDown : Bool;
      qConvRun_TTUp : Bool;
      qDelStprDown_TTUp : Bool;
      qOTS_Frm_TTDown : Bool;
      qOTS_Frm_TTUp : Bool;
      qOutput1 : Bool;
      qProcessStart : Bool;
      qRTR_Frm_TTDwn : Bool;
      qRTR_Frm_TTUp : Bool;
      qStprDown_TTDown : Bool;
      qStprDown_TTUp : Bool;
      qStprRaise_TTDown : Bool;
      qStprRaise_TTUp : Bool;
      qTTLockCmd : Bool;
      qTTUnlockCmd : Bool;
      qTT_0Deg : Bool;
      qTT_90Deg : Bool;
   END_VAR
   VAR_IN_OUT
      iqRX_Frn_Prev_TtDown : Bool;
      iqRx_Frm_Prev_TTUp : Bool;
      iqTx_To_Next_0DegTTDown : Bool;
      iqTx_To_Next_0DegTTUp : Bool;
      iqTx_To_Next_90DegTTUp : Bool;
   END_VAR
   VAR DB_SPECIFIC
      StateNo : Int;
      s100_StWtForTTUnlck : Bool;
      s100_StWtForTTUnlck_T1 : Bool;
      s10_StRecoveryCondition : Bool;
      s10_StRecoveryCondition_T1 : Bool;
      s10_StRecoveryCondition_T2 : Bool;
      s10_StRecoveryCondition_T3 : Bool;
      s10_StRecoveryCondition_T4 : Bool;
      s10_StRecoveryCondition_T5 : Bool;
      s10_StRecoveryCondition_T6 : Bool;
      s10_StRecoveryCondition_T7 : Bool;
      s110_StWtForTTTurn90 : Bool;
      s110_StWtForTTTurn90_T1 : Bool;
      s120_StWtForTTLck : Bool;
      s120_StWtForTTLck_T1 : Bool;
      s130_StChkTTDwnRdyToRecv : Bool;
      s130_StChkTTDwnRdyToRecv_T1 : Bool;
      s130_StChkTTDwnRdyToRecv_T2 : Bool;
      s140_StWtFrConveyorStrt : Bool;
      s140_StWtFrConveyorStrt_T1 : Bool;
      s150_StChkNxtStRdyToRecvTTUp : Bool;
      s150_StChkNxtStRdyToRecvTTUp_T1 : Bool;
      s150_StChkNxtStRdyToRecvTTUp_T2 : Bool;
      s15_StWaitForManCorrection : Bool;
      s15_StWaitForManCorrection_T1 : Bool;
      s160_StWtFrStprDn_CnvyrStrt : Bool;
      s160_StWtFrStprDn_CnvyrStrt_T1 : Bool;
      s165_StWtPalAbsnt : Bool;
      s165_StWtPalAbsnt_T1 : Bool;
      s167_StWtFrDeforkOvr : Bool;
      s167_StWtFrDeforkOvr_Cond1 : Bool;
      s167_StWtFrDeforkOvr_Cond2 : Bool;
      s167_StWtFrDeforkOvr_T1 : Bool;
      s170_StWtForTTUpStprUp : Bool;
      s170_StWtForTTUpStprUp_T1 : Bool;
      s180_StWtForTTUnlk : Bool;
      s180_StWtForTTUnlk_T1 : Bool;
      s190_StWtForTT_To_0 : Bool;
      s190_StWtForTT_To_0_T1 : Bool;
      s192_StWtForTTlok : Bool;
      s192_StWtForTTlok_T1 : Bool;
      s20_StChkForPalletPresent : Bool;
      s20_StChkForPalletPresent_T1 : Bool;
      s20_StChkForPalletPresent_T2 : Bool;
      s20_StChkForPalletPresent_T3 : Bool;
      s20_StChkForPalletPresent_T4 : Bool;
      s210_StWtFrTTUnlk : Bool;
      s210_StWtFrTTUnlk_T1 : Bool;
      s220_StWtFrTT_Trn_0 : Bool;
      s220_StWtFrTT_Trn_0_T1 : Bool;
      s230_StWtFrTTLock : Bool;
      s230_StWtFrTTLock_T1 : Bool;
      s240_StWtFRTRNxtStnTTDown : Bool;
      s240_StWtFRTRNxtStnTTDown_T1 : Bool;
      s240_StWtFRTRNxtStnTTDown_T2 : Bool;
      s250_StWtTTDnStprDn_CnvyrStr : Bool;
      s250_StWtTTDnStprDn_CnvyrStr_T1 : Bool;
      s260_StWtPalAbsent : Bool;
      s260_StWtPalAbsent_T1 : Bool;
      s270_StWtFrTTDwnStprUp : Bool;
      s270_StWtFrTTDwnStprUp_T1 : Bool;
      s280_StWtRFrOTSFRmPrev_TTUp : Bool;
      s280_StWtRFrOTSFRmPrev_TTUp_T1 : Bool;
      s290_StWtFrTTUpCnvyrStrt : Bool;
      s290_StWtFrTTUpCnvyrStrt_T1 : Bool;
      s300_StChkTTPos : Bool;
      s300_StChkTTPos_T1 : Bool;
      s300_StChkTTPos_T2 : Bool;
      s300_StChkTTPos_T3 : Bool;
      s30_StChckPartSts : Bool;
      s30_StChckPartSts_T1 : Bool;
      s310_StWtRTRFrmTTUpAt0 : Bool;
      s310_StWtRTRFrmTTUpAt0_T1 : Bool;
      s310_StWtRTRFrmTTUpAt0_T2 : Bool;
      s320_StWtFrTTUpCnvyrStrtAt0 : Bool;
      s320_StWtFrTTUpCnvyrStrtAt0_T1 : Bool;
      s340_StChkTTDwnRdyToRecvAt90 : Bool;
      s340_StChkTTDwnRdyToRecvAt90_T1 : Bool;
      s340_StChkTTDwnRdyToRecvAt90_T2 : Bool;
      s350_StWtCnvyrStrt90 : Bool;
      s350_StWtCnvyrStrt90_T1 : Bool;
      s365_StWtForTTUlkAtIbtwn : Bool;
      s365_StWtForTTUlkAtIbtwn_T1 : Bool;
      s370_StWtForTTTurnZrAtIbtwn : Bool;
      s370_StWtForTTTurnZrAtIbtwn_T1 : Bool;
      s380_StWtForTTLock : Bool;
      s380_StWtForTTLock_T1 : Bool;
      s400_StWt2Defork : Bool;
      s400_StWt2Defork_Cond1 : Bool;
      s400_StWt2Defork_Cond2 : Bool;
      s400_StWt2Defork_T1 : Bool;
      s40_StWtForTTUnlock : Bool;
      s40_StWtForTTUnlock_T1 : Bool;
      s410_StWtForTTUlkAtIbtwn : Bool;
      s410_StWtForTTUlkAtIbtwn_T1 : Bool;
      s415_StWtForTTTurn90AtIbtwn : Bool;
      s415_StWtForTTTurn90AtIbtwn_T1 : Bool;
      s420_StWtForTTLock1 : Bool;
      s420_StWtForTTLock1_T1 : Bool;
      s50_StWtForTTTurn0 : Bool;
      s50_StWtForTTTurn0_T1 : Bool;
      s60_StWtForTTLock : Bool;
      s60_StWtForTTLock_T1 : Bool;
      s70_StWtOTSfrmTTUp : Bool;
      s70_StWtOTSfrmTTUp_T1 : Bool;
      s80_StWtTTUpStpDwnCnvrStrt : Bool;
      s80_StWtTTUpStpDwnCnvrStrt_T1 : Bool;
      s85_StWtPalPresntAtRej : Bool;
      s85_StWtPalPresntAtRej_T1 : Bool;
      s90_StWtTTUpStprUp : Bool;
      s90_StWtTTUpStprUp_T1 : Bool;
      sDefork1Done : Bool;
      sDefork2Done : Bool;
      sOTSFrmDwnTout : Bool;
      sOTSFrmUpTout : Bool;
      sPalOnStop_TTDown : Bool;
      sPalOnStop_TTUp_0Deg : Bool;
      sPalOnStop_TTUp_90Deg : Bool;
      sPalletAbsnDebTTUp : Bool;
      sPalletAbsntDebTTDown : Bool;
      sPalletAbsntDebTTUp : Bool;
      sPalletPrsntDebTTDown : Bool;
      sPalletPrsntDebTTUp : Bool;
      sRTRFrmUpTout : Bool;
      sSst : Bool;
      sSstPulse : Bool;
      sSstRise : Bool;
      sStWtResetRel : Bool;
      sStWtResetRel_T1 : Bool;
      sTTDwnSeqOver : Bool;
      sTTDwn_0Pos_TX_Time : Bool;
      sTTDwn_90Pos_RX_Time : Bool;
      sTTDwn_Timer_ON : Bool;
      sTTUpSeqOver : Bool;
      sTTUp_90Pos_TX_Time : Bool;
      sTTUp_Timer_ON : Bool;
      sTrBothPalletPresent : Bool;
   END_VAR
   VAR_TEMP
      tOne : Bool;
   END_VAR
   VAR_TEMP   // added for the SCL form of the ladder/FBD networks
      _w1 : Bool;
   END_VAR
BEGIN

REGION Network 1
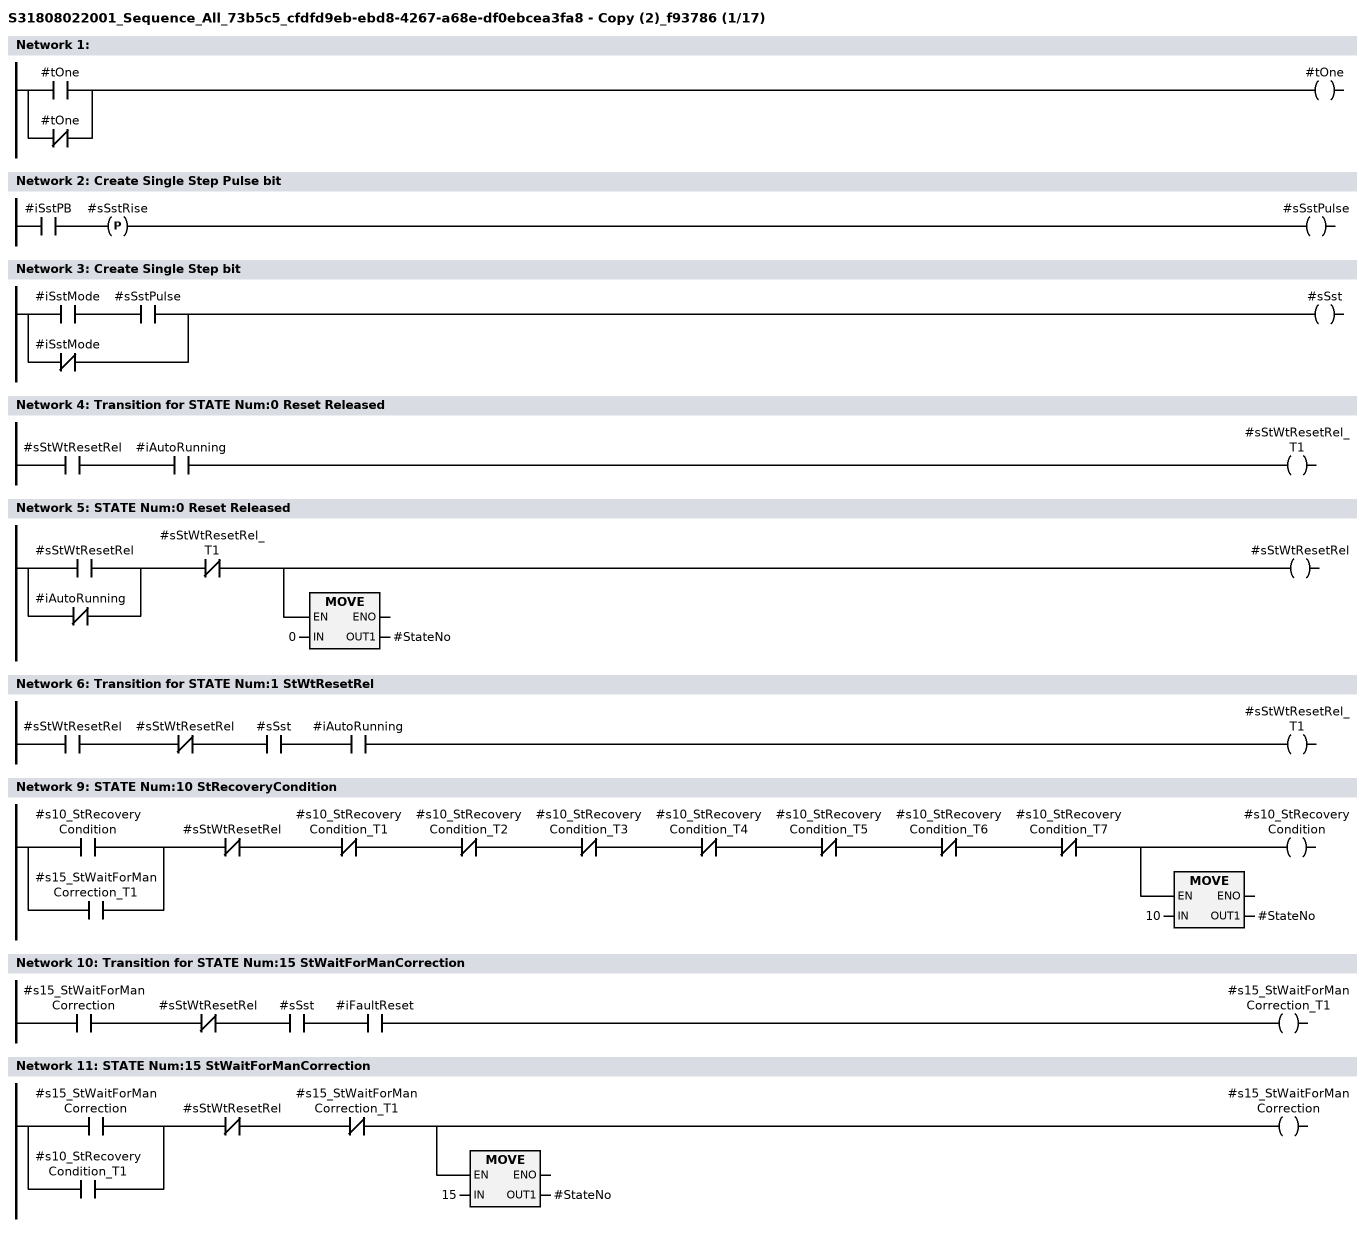
   RUNG wire#powerrail
      Contact( #tOne )
      wire#w1
      Coil( #tOne )
   END_RUNG
   RUNG wire#powerrail
      I_Contact( #tOne )
   END_RUNG wire#w1
   // the same network as SCL:
   #tOne := #tOne OR NOT #tOne;
END_REGION

REGION Network 2: Create Single Step Pulse bit
   RUNG wire#powerrail
      Contact( #iSstPB )
      P_Trig( #sSstRise )
      Coil( #sSstPulse )
   END_RUNG
   // the same network as SCL:
   #_w1 := #iSstPB AND NOT #sSstRise;   // rising edge
   #sSstRise := #iSstPB;
   #sSstPulse := #_w1;
END_REGION

REGION Network 3: Create Single Step bit
   RUNG wire#powerrail
      Contact( #iSstMode )
      Contact( #sSstPulse )
      wire#w1
      Coil( #sSst )
   END_RUNG
   RUNG wire#powerrail
      I_Contact( #iSstMode )
   END_RUNG wire#w1
   // the same network as SCL:
   #sSst := (#iSstMode AND #sSstPulse) OR NOT #iSstMode;
END_REGION

REGION Network 4: Transition for STATE Num:0 Reset Released
   RUNG wire#powerrail
      Contact( #sStWtResetRel )
      Contact( #iAutoRunning )
      Coil( #sStWtResetRel_T1 )
   END_RUNG
   // the same network as SCL:
   #sStWtResetRel_T1 := #sStWtResetRel AND #iAutoRunning;
END_REGION

REGION Network 5: STATE Num:0 Reset Released
   RUNG wire#powerrail
      Contact( #sStWtResetRel )
      wire#w1
      I_Contact( #sStWtResetRel_T1 )
      wire#w2
      Coil( #sStWtResetRel )
   END_RUNG
   RUNG wire#powerrail
      I_Contact( #iAutoRunning )
   END_RUNG wire#w1
   RUNG wire#w2
      { S7_GenerateENO := "TRUE" } Move(in := 0, out1 => #StateNo)
   END_RUNG
   // the same network as SCL:
   #sStWtResetRel := (#sStWtResetRel OR NOT #iAutoRunning) AND NOT #sStWtResetRel_T1;
   IF #sStWtResetRel THEN #StateNo := 0; END_IF;
END_REGION

REGION Network 6: Transition for STATE Num:1 StWtResetRel
   RUNG wire#powerrail
      Contact( #sStWtResetRel )
      I_Contact( #sStWtResetRel )
      Contact( #sSst )
      Contact( #iAutoRunning )
      Coil( #sStWtResetRel_T1 )
   END_RUNG
   // the same network as SCL:
   #sStWtResetRel_T1 := #sStWtResetRel AND NOT #sStWtResetRel AND #sSst AND #iAutoRunning;
END_REGION

NETWORK
TITLE = STATE Num:1 StWtResetRel
      A(;
      O     #sStWtResetRel;
//wrong transition variable removed
      );
      AN    #sStWtResetRel;
      AN    #sStWtResetRel_T1;
      =     %L1.0;
      A     %L1.0;
      BLD   102;
      =     #sStWtResetRel;
      A     %L1.0;
      JNB   Label_1;
      L     1;
      T     #StateNo;
Label_1:NOP   0;

NETWORK
TITLE = Transition for STATE Num:10 StRecoveryCondition
      A     #s10_StRecoveryCondition;
      AN    #sStWtResetRel;
      A     #sSst;
      =     %L1.0;
      A     %L1.0;
      A(;
      O(;
      A     #iRx_Frm_Prev_TTUp;
      AN    #iTTAt0Pos;
      );
      O(;
      A     #iqRX_Frn_Prev_TtDown;
      AN    #iTTAt90Pos;
      );
      O(;
      O     #iqTx_To_Next_90DegTTUp;
      O     #sPalOnStop_TTUp_90Deg;
      AN    #iTTAt90Pos;
      );
      O(;
      O     #iqTx_To_Next_0DegTTUp;
      O     #sPalOnStop_TTUp_0Deg;
      AN    #iTTAt0Pos;
      );
      O(;
      O     #iqTx_To_Next_0DegTTDown;
      O     #sPalOnStop_TTDown;
      AN    #iTTAt0Pos;
      );
      O(;
      O     #sPalOnStop_TTUp_0Deg;
      O     #sPalOnStop_TTUp_90Deg;
      O     #sPalOnStop_TTDown;
      A     #iTTUnlocked;
      );
      );
      =     #s10_StRecoveryCondition_T1;
      A     %L1.0;
      AN    #s10_StRecoveryCondition_T1;
      A(;
      O     #iqTx_To_Next_0DegTTUp;
      O     #sPalOnStop_TTUp_0Deg;
      );
      A     #iTTAt0Pos;
      A     #iTTLocked;
      =     #s10_StRecoveryCondition_T2;
      A     %L1.0;
      AN    #s10_StRecoveryCondition_T1;
      AN    #s10_StRecoveryCondition_T2;
      A(;
      O     #iqTx_To_Next_90DegTTUp;
      O     #sPalOnStop_TTUp_90Deg;
      );
      A     #iTTAt90Pos;
      A     #iTTLocked;
      =     #s10_StRecoveryCondition_T3;
      A     %L1.0;
      AN    #s10_StRecoveryCondition_T1;
      AN    #s10_StRecoveryCondition_T2;
      AN    #s10_StRecoveryCondition_T3;
      A(;
      O     #iqTx_To_Next_0DegTTDown;
      O     #sPalOnStop_TTDown;
      );
      A     #iTTAt0Pos;
      A     #iTTLocked;
      =     #s10_StRecoveryCondition_T4;
      A     %L1.0;
      AN    #s10_StRecoveryCondition_T1;
      AN    #s10_StRecoveryCondition_T2;
      AN    #s10_StRecoveryCondition_T3;
      AN    #s10_StRecoveryCondition_T4;
      A(;
      O     #iRx_Frm_Prev_TTUp;
      O     #iRecvAreaClr_TTUp;
      );
      A     #iTTAt0Pos;
      A     #iTTLocked;
      =     #s10_StRecoveryCondition_T5;
      A     %L1.0;
      AN    #s10_StRecoveryCondition_T1;
      AN    #s10_StRecoveryCondition_T2;
      AN    #s10_StRecoveryCondition_T3;
      AN    #s10_StRecoveryCondition_T4;
      AN    #s10_StRecoveryCondition_T5;
      A(;
      O     #iqRX_Frn_Prev_TtDown;
      ON    #iRecvAreaClr_TTDown;
      );
      A     #iTTAt90Pos;
      A     #iTTLocked;
      =     #s10_StRecoveryCondition_T6;
      A     %L1.0;
      AN    #s10_StRecoveryCondition_T1;
      AN    #s10_StRecoveryCondition_T2;
      AN    #s10_StRecoveryCondition_T3;
      AN    #s10_StRecoveryCondition_T4;
      AN    #s10_StRecoveryCondition_T5;
      AN    #s10_StRecoveryCondition_T6;
      A(;
      A(;
      A     #iXferAreaClr_90DegTTUp;
      A     #iXferAreaClr_0DegTTDown;
      A     #iRecvAreaClr_TTDown;
      A     #iRecvAreaClr_TTUp;
      );
      O(;
      AN    #sPalOnStop_TTUp_0Deg;
      AN    #sPalOnStop_TTUp_90Deg;
      AN    #sPalOnStop_TTDown;
      );
      O(;
      AN    #iqTx_To_Next_90DegTTUp;
      AN    #iqTx_To_Next_0DegTTUp;
      AN    #iqTx_To_Next_0DegTTDown;
      AN    #iqRX_Frn_Prev_TtDown;
      AN    #iRx_Frm_Prev_TTUp;
      );
      );
      =     #s10_StRecoveryCondition_T7;

REGION Network 9: STATE Num:10 StRecoveryCondition
   RUNG wire#powerrail
      Contact( #s10_StRecoveryCondition )
      wire#w1
      I_Contact( #sStWtResetRel )
      I_Contact( #s10_StRecoveryCondition_T1 )
      I_Contact( #s10_StRecoveryCondition_T2 )
      I_Contact( #s10_StRecoveryCondition_T3 )
      I_Contact( #s10_StRecoveryCondition_T4 )
      I_Contact( #s10_StRecoveryCondition_T5 )
      I_Contact( #s10_StRecoveryCondition_T6 )
      I_Contact( #s10_StRecoveryCondition_T7 )
      wire#w2
      Coil( #s10_StRecoveryCondition )
   END_RUNG
   RUNG wire#powerrail
      Contact( #s15_StWaitForManCorrection_T1 )
   END_RUNG wire#w1
   RUNG wire#w2
      { S7_GenerateENO := "TRUE" } Move(in := 10, out1 => #StateNo)
   END_RUNG
   // the same network as SCL:
   #s10_StRecoveryCondition := (#s10_StRecoveryCondition OR #s15_StWaitForManCorrection_T1) AND NOT #sStWtResetRel AND NOT #s10_StRecoveryCondition_T1 AND NOT #s10_StRecoveryCondition_T2 AND NOT #s10_StRecoveryCondition_T3 AND NOT #s10_StRecoveryCondition_T4 AND NOT #s10_StRecoveryCondition_T5 AND NOT #s10_StRecoveryCondition_T6 AND NOT #s10_StRecoveryCondition_T7;
   IF #s10_StRecoveryCondition THEN #StateNo := 10; END_IF;
END_REGION

REGION Network 10: Transition for STATE Num:15 StWaitForManCorrection
   RUNG wire#powerrail
      Contact( #s15_StWaitForManCorrection )
      I_Contact( #sStWtResetRel )
      Contact( #sSst )
      Contact( #iFaultReset )
      Coil( #s15_StWaitForManCorrection_T1 )
   END_RUNG
   // the same network as SCL:
   #s15_StWaitForManCorrection_T1 := #s15_StWaitForManCorrection AND NOT #sStWtResetRel AND #sSst AND #iFaultReset;
END_REGION

REGION Network 11: STATE Num:15 StWaitForManCorrection
   RUNG wire#powerrail
      Contact( #s15_StWaitForManCorrection )
      wire#w1
      I_Contact( #sStWtResetRel )
      I_Contact( #s15_StWaitForManCorrection_T1 )
      wire#w2
      Coil( #s15_StWaitForManCorrection )
   END_RUNG
   RUNG wire#powerrail
      Contact( #s10_StRecoveryCondition_T1 )
   END_RUNG wire#w1
   RUNG wire#w2
      { S7_GenerateENO := "TRUE" } Move(in := 15, out1 => #StateNo)
   END_RUNG
   // the same network as SCL:
   #s15_StWaitForManCorrection := (#s15_StWaitForManCorrection OR #s10_StRecoveryCondition_T1) AND NOT #sStWtResetRel AND NOT #s15_StWaitForManCorrection_T1;
   IF #s15_StWaitForManCorrection THEN #StateNo := 15; END_IF;
END_REGION

REGION Network 12: Transition for STATE Num:20 StChkForPalletPresent
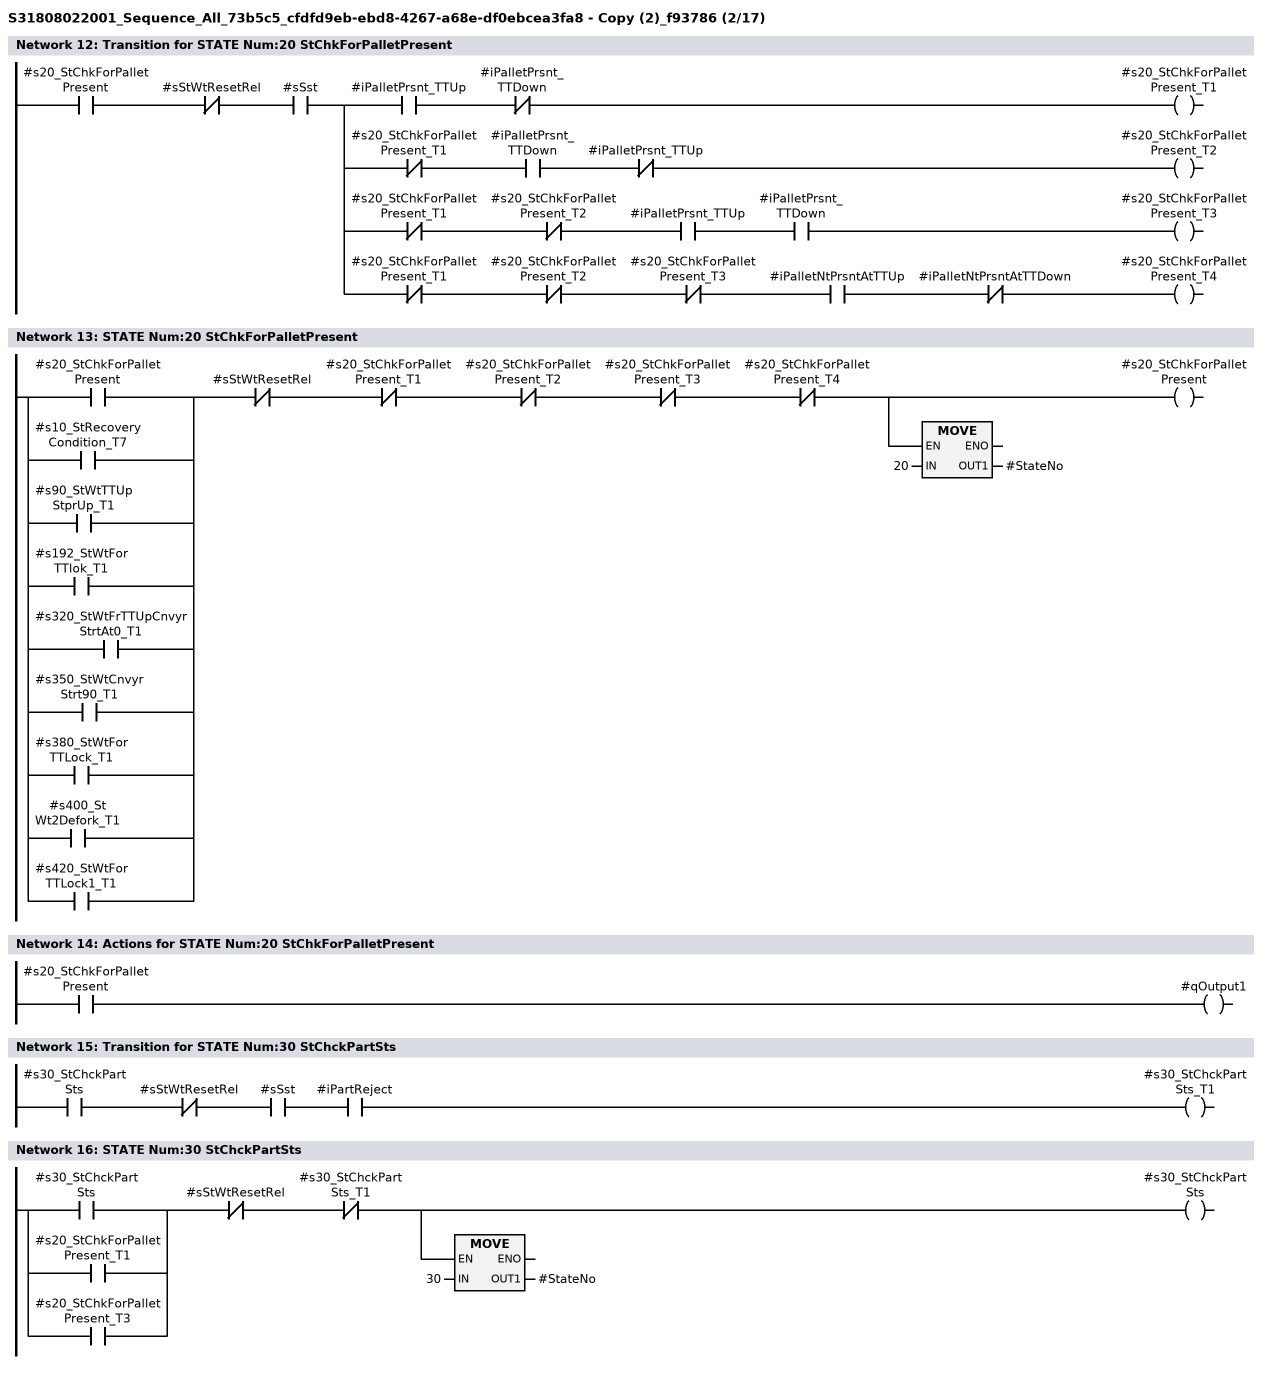
   RUNG wire#powerrail
      Contact( #s20_StChkForPalletPresent )
      I_Contact( #sStWtResetRel )
      Contact( #sSst )
      wire#w1
      Contact( #iPalletPrsnt_TTUp )
      I_Contact( #iPalletPrsnt_TTDown )
      Coil( #s20_StChkForPalletPresent_T1 )
   END_RUNG
   RUNG wire#w1
      I_Contact( #s20_StChkForPalletPresent_T1 )
      Contact( #iPalletPrsnt_TTDown )
      I_Contact( #iPalletPrsnt_TTUp )
      Coil( #s20_StChkForPalletPresent_T2 )
   END_RUNG
   RUNG wire#w1
      I_Contact( #s20_StChkForPalletPresent_T1 )
      I_Contact( #s20_StChkForPalletPresent_T2 )
      Contact( #iPalletPrsnt_TTUp )
      Contact( #iPalletPrsnt_TTDown )
      Coil( #s20_StChkForPalletPresent_T3 )
   END_RUNG
   RUNG wire#w1
      I_Contact( #s20_StChkForPalletPresent_T1 )
      I_Contact( #s20_StChkForPalletPresent_T2 )
      I_Contact( #s20_StChkForPalletPresent_T3 )
      Contact( #iPalletNtPrsntAtTTUp )
      I_Contact( #iPalletNtPrsntAtTTDown )
      Coil( #s20_StChkForPalletPresent_T4 )
   END_RUNG
   // the same network as SCL:
   #_w1 := #s20_StChkForPalletPresent AND NOT #sStWtResetRel AND #sSst;
   #s20_StChkForPalletPresent_T1 := #_w1 AND #iPalletPrsnt_TTUp AND NOT #iPalletPrsnt_TTDown;
   #s20_StChkForPalletPresent_T2 := #_w1 AND NOT #s20_StChkForPalletPresent_T1 AND #iPalletPrsnt_TTDown AND NOT #iPalletPrsnt_TTUp;
   #s20_StChkForPalletPresent_T3 := #_w1 AND NOT #s20_StChkForPalletPresent_T1 AND NOT #s20_StChkForPalletPresent_T2 AND #iPalletPrsnt_TTUp AND #iPalletPrsnt_TTDown;
   #s20_StChkForPalletPresent_T4 := #_w1 AND NOT #s20_StChkForPalletPresent_T1 AND NOT #s20_StChkForPalletPresent_T2 AND NOT #s20_StChkForPalletPresent_T3 AND #iPalletNtPrsntAtTTUp AND NOT #iPalletNtPrsntAtTTDown;
END_REGION

REGION Network 13: STATE Num:20 StChkForPalletPresent
   RUNG wire#powerrail
      Contact( #s20_StChkForPalletPresent )
      wire#w1
      I_Contact( #sStWtResetRel )
      I_Contact( #s20_StChkForPalletPresent_T1 )
      I_Contact( #s20_StChkForPalletPresent_T2 )
      I_Contact( #s20_StChkForPalletPresent_T3 )
      I_Contact( #s20_StChkForPalletPresent_T4 )
      wire#w2
      Coil( #s20_StChkForPalletPresent )
   END_RUNG
   RUNG wire#powerrail
      Contact( #s10_StRecoveryCondition_T7 )
   END_RUNG wire#w1
   RUNG wire#powerrail
      Contact( #s90_StWtTTUpStprUp_T1 )
   END_RUNG wire#w1
   RUNG wire#powerrail
      Contact( #s192_StWtForTTlok_T1 )
   END_RUNG wire#w1
   RUNG wire#powerrail
      Contact( #s320_StWtFrTTUpCnvyrStrtAt0_T1 )
   END_RUNG wire#w1
   RUNG wire#powerrail
      Contact( #s350_StWtCnvyrStrt90_T1 )
   END_RUNG wire#w1
   RUNG wire#powerrail
      Contact( #s380_StWtForTTLock_T1 )
   END_RUNG wire#w1
   RUNG wire#powerrail
      Contact( #s400_StWt2Defork_T1 )
   END_RUNG wire#w1
   RUNG wire#powerrail
      Contact( #s420_StWtForTTLock1_T1 )
   END_RUNG wire#w1
   RUNG wire#w2
      { S7_GenerateENO := "TRUE" } Move(in := 20, out1 => #StateNo)
   END_RUNG
   // the same network as SCL:
   #s20_StChkForPalletPresent := (#s20_StChkForPalletPresent OR #s10_StRecoveryCondition_T7 OR #s90_StWtTTUpStprUp_T1 OR #s192_StWtForTTlok_T1 OR #s320_StWtFrTTUpCnvyrStrtAt0_T1 OR #s350_StWtCnvyrStrt90_T1 OR #s380_StWtForTTLock_T1 OR #s400_StWt2Defork_T1 OR #s420_StWtForTTLock1_T1) AND NOT #sStWtResetRel AND NOT #s20_StChkForPalletPresent_T1 AND NOT #s20_StChkForPalletPresent_T2 AND NOT #s20_StChkForPalletPresent_T3 AND NOT #s20_StChkForPalletPresent_T4;
   IF #s20_StChkForPalletPresent THEN #StateNo := 20; END_IF;
END_REGION

REGION Network 14: Actions for STATE Num:20 StChkForPalletPresent
   RUNG wire#powerrail
      Contact( #s20_StChkForPalletPresent )
      Coil( #qOutput1 )
   END_RUNG
   // the same network as SCL:
   #qOutput1 := #s20_StChkForPalletPresent;
END_REGION

REGION Network 15: Transition for STATE Num:30 StChckPartSts
   RUNG wire#powerrail
      Contact( #s30_StChckPartSts )
      I_Contact( #sStWtResetRel )
      Contact( #sSst )
      Contact( #iPartReject )
      Coil( #s30_StChckPartSts_T1 )
   END_RUNG
   // the same network as SCL:
   #s30_StChckPartSts_T1 := #s30_StChckPartSts AND NOT #sStWtResetRel AND #sSst AND #iPartReject;
END_REGION

REGION Network 16: STATE Num:30 StChckPartSts
   RUNG wire#powerrail
      Contact( #s30_StChckPartSts )
      wire#w1
      I_Contact( #sStWtResetRel )
      I_Contact( #s30_StChckPartSts_T1 )
      wire#w2
      Coil( #s30_StChckPartSts )
   END_RUNG
   RUNG wire#powerrail
      Contact( #s20_StChkForPalletPresent_T1 )
   END_RUNG wire#w1
   RUNG wire#powerrail
      Contact( #s20_StChkForPalletPresent_T3 )
   END_RUNG wire#w1
   RUNG wire#w2
      { S7_GenerateENO := "TRUE" } Move(in := 30, out1 => #StateNo)
   END_RUNG
   // the same network as SCL:
   #s30_StChckPartSts := (#s30_StChckPartSts OR #s20_StChkForPalletPresent_T1 OR #s20_StChkForPalletPresent_T3) AND NOT #sStWtResetRel AND NOT #s30_StChckPartSts_T1;
   IF #s30_StChckPartSts THEN #StateNo := 30; END_IF;
END_REGION

REGION Network 17: Actions for STATE Num:30 StChckPartSts
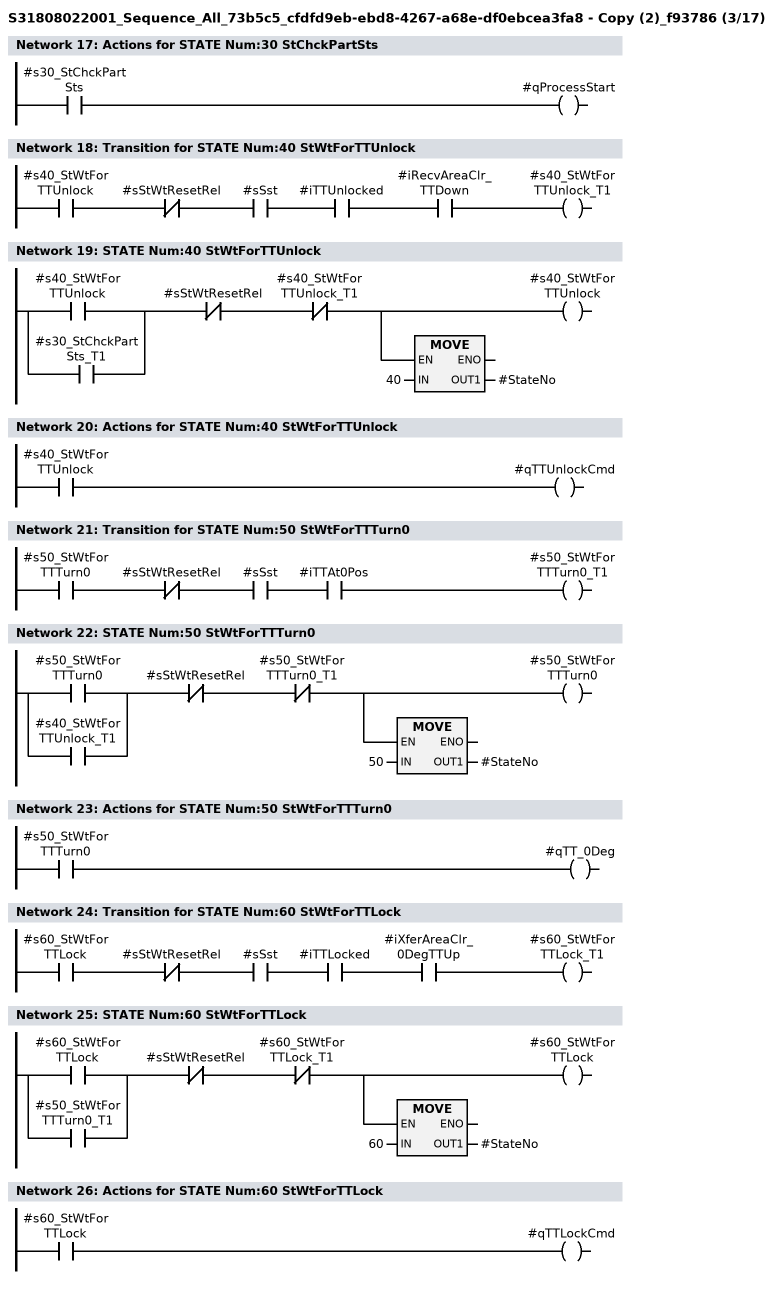
   RUNG wire#powerrail
      Contact( #s30_StChckPartSts )
      Coil( #qProcessStart )
   END_RUNG
   // the same network as SCL:
   #qProcessStart := #s30_StChckPartSts;
END_REGION

REGION Network 18: Transition for STATE Num:40 StWtForTTUnlock
   RUNG wire#powerrail
      Contact( #s40_StWtForTTUnlock )
      I_Contact( #sStWtResetRel )
      Contact( #sSst )
      Contact( #iTTUnlocked )
      Contact( #iRecvAreaClr_TTDown )
      Coil( #s40_StWtForTTUnlock_T1 )
   END_RUNG
   // the same network as SCL:
   #s40_StWtForTTUnlock_T1 := #s40_StWtForTTUnlock AND NOT #sStWtResetRel AND #sSst AND #iTTUnlocked AND #iRecvAreaClr_TTDown;
END_REGION

REGION Network 19: STATE Num:40 StWtForTTUnlock
   RUNG wire#powerrail
      Contact( #s40_StWtForTTUnlock )
      wire#w1
      I_Contact( #sStWtResetRel )
      I_Contact( #s40_StWtForTTUnlock_T1 )
      wire#w2
      Coil( #s40_StWtForTTUnlock )
   END_RUNG
   RUNG wire#powerrail
      Contact( #s30_StChckPartSts_T1 )
   END_RUNG wire#w1
   RUNG wire#w2
      { S7_GenerateENO := "TRUE" } Move(in := 40, out1 => #StateNo)
   END_RUNG
   // the same network as SCL:
   #s40_StWtForTTUnlock := (#s40_StWtForTTUnlock OR #s30_StChckPartSts_T1) AND NOT #sStWtResetRel AND NOT #s40_StWtForTTUnlock_T1;
   IF #s40_StWtForTTUnlock THEN #StateNo := 40; END_IF;
END_REGION

REGION Network 20: Actions for STATE Num:40 StWtForTTUnlock
   RUNG wire#powerrail
      Contact( #s40_StWtForTTUnlock )
      Coil( #qTTUnlockCmd )
   END_RUNG
   // the same network as SCL:
   #qTTUnlockCmd := #s40_StWtForTTUnlock;
END_REGION

REGION Network 21: Transition for STATE Num:50 StWtForTTTurn0
   RUNG wire#powerrail
      Contact( #s50_StWtForTTTurn0 )
      I_Contact( #sStWtResetRel )
      Contact( #sSst )
      Contact( #iTTAt0Pos )
      Coil( #s50_StWtForTTTurn0_T1 )
   END_RUNG
   // the same network as SCL:
   #s50_StWtForTTTurn0_T1 := #s50_StWtForTTTurn0 AND NOT #sStWtResetRel AND #sSst AND #iTTAt0Pos;
END_REGION

REGION Network 22: STATE Num:50 StWtForTTTurn0
   RUNG wire#powerrail
      Contact( #s50_StWtForTTTurn0 )
      wire#w1
      I_Contact( #sStWtResetRel )
      I_Contact( #s50_StWtForTTTurn0_T1 )
      wire#w2
      Coil( #s50_StWtForTTTurn0 )
   END_RUNG
   RUNG wire#powerrail
      Contact( #s40_StWtForTTUnlock_T1 )
   END_RUNG wire#w1
   RUNG wire#w2
      { S7_GenerateENO := "TRUE" } Move(in := 50, out1 => #StateNo)
   END_RUNG
   // the same network as SCL:
   #s50_StWtForTTTurn0 := (#s50_StWtForTTTurn0 OR #s40_StWtForTTUnlock_T1) AND NOT #sStWtResetRel AND NOT #s50_StWtForTTTurn0_T1;
   IF #s50_StWtForTTTurn0 THEN #StateNo := 50; END_IF;
END_REGION

REGION Network 23: Actions for STATE Num:50 StWtForTTTurn0
   RUNG wire#powerrail
      Contact( #s50_StWtForTTTurn0 )
      Coil( #qTT_0Deg )
   END_RUNG
   // the same network as SCL:
   #qTT_0Deg := #s50_StWtForTTTurn0;
END_REGION

REGION Network 24: Transition for STATE Num:60 StWtForTTLock
   RUNG wire#powerrail
      Contact( #s60_StWtForTTLock )
      I_Contact( #sStWtResetRel )
      Contact( #sSst )
      Contact( #iTTLocked )
      Contact( #iXferAreaClr_0DegTTUp )
      Coil( #s60_StWtForTTLock_T1 )
   END_RUNG
   // the same network as SCL:
   #s60_StWtForTTLock_T1 := #s60_StWtForTTLock AND NOT #sStWtResetRel AND #sSst AND #iTTLocked AND #iXferAreaClr_0DegTTUp;
END_REGION

REGION Network 25: STATE Num:60 StWtForTTLock
   RUNG wire#powerrail
      Contact( #s60_StWtForTTLock )
      wire#w1
      I_Contact( #sStWtResetRel )
      I_Contact( #s60_StWtForTTLock_T1 )
      wire#w2
      Coil( #s60_StWtForTTLock )
   END_RUNG
   RUNG wire#powerrail
      Contact( #s50_StWtForTTTurn0_T1 )
   END_RUNG wire#w1
   RUNG wire#w2
      { S7_GenerateENO := "TRUE" } Move(in := 60, out1 => #StateNo)
   END_RUNG
   // the same network as SCL:
   #s60_StWtForTTLock := (#s60_StWtForTTLock OR #s50_StWtForTTTurn0_T1) AND NOT #sStWtResetRel AND NOT #s60_StWtForTTLock_T1;
   IF #s60_StWtForTTLock THEN #StateNo := 60; END_IF;
END_REGION

REGION Network 26: Actions for STATE Num:60 StWtForTTLock
   RUNG wire#powerrail
      Contact( #s60_StWtForTTLock )
      Coil( #qTTLockCmd )
   END_RUNG
   // the same network as SCL:
   #qTTLockCmd := #s60_StWtForTTLock;
END_REGION

REGION Network 27: Transition for STATE Num:70 StWtOTSfrmTTUp
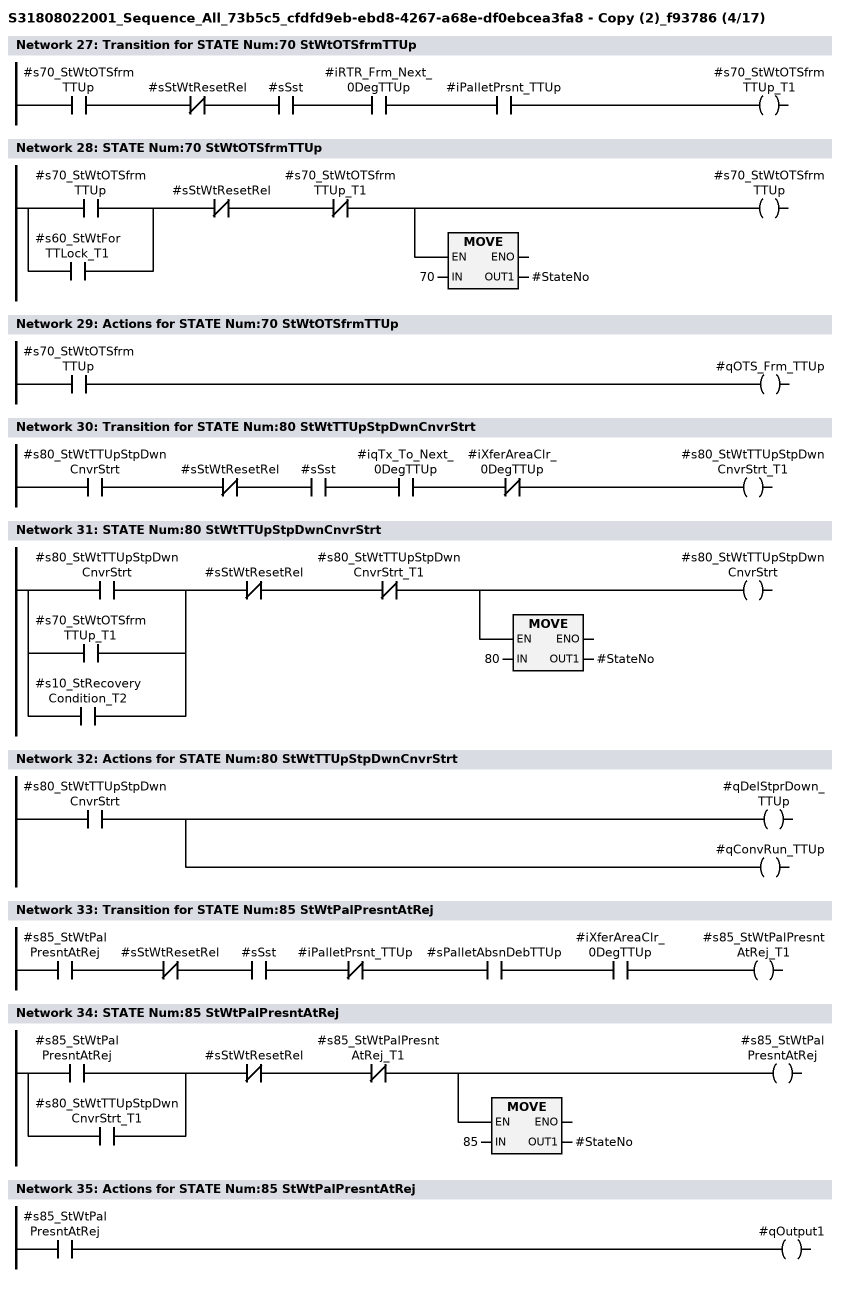
   RUNG wire#powerrail
      Contact( #s70_StWtOTSfrmTTUp )
      I_Contact( #sStWtResetRel )
      Contact( #sSst )
      Contact( #iRTR_Frm_Next_0DegTTUp )
      Contact( #iPalletPrsnt_TTUp )
      Coil( #s70_StWtOTSfrmTTUp_T1 )
   END_RUNG
   // the same network as SCL:
   #s70_StWtOTSfrmTTUp_T1 := #s70_StWtOTSfrmTTUp AND NOT #sStWtResetRel AND #sSst AND #iRTR_Frm_Next_0DegTTUp AND #iPalletPrsnt_TTUp;
END_REGION

REGION Network 28: STATE Num:70 StWtOTSfrmTTUp
   RUNG wire#powerrail
      Contact( #s70_StWtOTSfrmTTUp )
      wire#w1
      I_Contact( #sStWtResetRel )
      I_Contact( #s70_StWtOTSfrmTTUp_T1 )
      wire#w2
      Coil( #s70_StWtOTSfrmTTUp )
   END_RUNG
   RUNG wire#powerrail
      Contact( #s60_StWtForTTLock_T1 )
   END_RUNG wire#w1
   RUNG wire#w2
      { S7_GenerateENO := "TRUE" } Move(in := 70, out1 => #StateNo)
   END_RUNG
   // the same network as SCL:
   #s70_StWtOTSfrmTTUp := (#s70_StWtOTSfrmTTUp OR #s60_StWtForTTLock_T1) AND NOT #sStWtResetRel AND NOT #s70_StWtOTSfrmTTUp_T1;
   IF #s70_StWtOTSfrmTTUp THEN #StateNo := 70; END_IF;
END_REGION

REGION Network 29: Actions for STATE Num:70 StWtOTSfrmTTUp
   RUNG wire#powerrail
      Contact( #s70_StWtOTSfrmTTUp )
      Coil( #qOTS_Frm_TTUp )
   END_RUNG
   // the same network as SCL:
   #qOTS_Frm_TTUp := #s70_StWtOTSfrmTTUp;
END_REGION

REGION Network 30: Transition for STATE Num:80 StWtTTUpStpDwnCnvrStrt
   RUNG wire#powerrail
      Contact( #s80_StWtTTUpStpDwnCnvrStrt )
      I_Contact( #sStWtResetRel )
      Contact( #sSst )
      Contact( #iqTx_To_Next_0DegTTUp )
      I_Contact( #iXferAreaClr_0DegTTUp )
      Coil( #s80_StWtTTUpStpDwnCnvrStrt_T1 )
   END_RUNG
   // the same network as SCL:
   #s80_StWtTTUpStpDwnCnvrStrt_T1 := #s80_StWtTTUpStpDwnCnvrStrt AND NOT #sStWtResetRel AND #sSst AND #iqTx_To_Next_0DegTTUp AND NOT #iXferAreaClr_0DegTTUp;
END_REGION

REGION Network 31: STATE Num:80 StWtTTUpStpDwnCnvrStrt
   RUNG wire#powerrail
      Contact( #s80_StWtTTUpStpDwnCnvrStrt )
      wire#w1
      I_Contact( #sStWtResetRel )
      I_Contact( #s80_StWtTTUpStpDwnCnvrStrt_T1 )
      wire#w2
      Coil( #s80_StWtTTUpStpDwnCnvrStrt )
   END_RUNG
   RUNG wire#powerrail
      Contact( #s70_StWtOTSfrmTTUp_T1 )
   END_RUNG wire#w1
   RUNG wire#powerrail
      Contact( #s10_StRecoveryCondition_T2 )
   END_RUNG wire#w1
   RUNG wire#w2
      { S7_GenerateENO := "TRUE" } Move(in := 80, out1 => #StateNo)
   END_RUNG
   // the same network as SCL:
   #s80_StWtTTUpStpDwnCnvrStrt := (#s80_StWtTTUpStpDwnCnvrStrt OR #s70_StWtOTSfrmTTUp_T1 OR #s10_StRecoveryCondition_T2) AND NOT #sStWtResetRel AND NOT #s80_StWtTTUpStpDwnCnvrStrt_T1;
   IF #s80_StWtTTUpStpDwnCnvrStrt THEN #StateNo := 80; END_IF;
END_REGION

REGION Network 32: Actions for STATE Num:80 StWtTTUpStpDwnCnvrStrt
   RUNG wire#powerrail
      Contact( #s80_StWtTTUpStpDwnCnvrStrt )
      wire#w1
      Coil( #qDelStprDown_TTUp )
   END_RUNG
   RUNG wire#w1
      Coil( #qConvRun_TTUp )
   END_RUNG
   // the same network as SCL:
   #qDelStprDown_TTUp := #s80_StWtTTUpStpDwnCnvrStrt;
   #qConvRun_TTUp := #s80_StWtTTUpStpDwnCnvrStrt;
END_REGION

REGION Network 33: Transition for STATE Num:85 StWtPalPresntAtRej
   RUNG wire#powerrail
      Contact( #s85_StWtPalPresntAtRej )
      I_Contact( #sStWtResetRel )
      Contact( #sSst )
      I_Contact( #iPalletPrsnt_TTUp )
      Contact( #sPalletAbsnDebTTUp )
      Contact( #iXferAreaClr_0DegTTUp )
      Coil( #s85_StWtPalPresntAtRej_T1 )
   END_RUNG
   // the same network as SCL:
   #s85_StWtPalPresntAtRej_T1 := #s85_StWtPalPresntAtRej AND NOT #sStWtResetRel AND #sSst AND NOT #iPalletPrsnt_TTUp AND #sPalletAbsnDebTTUp AND #iXferAreaClr_0DegTTUp;
END_REGION

REGION Network 34: STATE Num:85 StWtPalPresntAtRej
   RUNG wire#powerrail
      Contact( #s85_StWtPalPresntAtRej )
      wire#w1
      I_Contact( #sStWtResetRel )
      I_Contact( #s85_StWtPalPresntAtRej_T1 )
      wire#w2
      Coil( #s85_StWtPalPresntAtRej )
   END_RUNG
   RUNG wire#powerrail
      Contact( #s80_StWtTTUpStpDwnCnvrStrt_T1 )
   END_RUNG wire#w1
   RUNG wire#w2
      { S7_GenerateENO := "TRUE" } Move(in := 85, out1 => #StateNo)
   END_RUNG
   // the same network as SCL:
   #s85_StWtPalPresntAtRej := (#s85_StWtPalPresntAtRej OR #s80_StWtTTUpStpDwnCnvrStrt_T1) AND NOT #sStWtResetRel AND NOT #s85_StWtPalPresntAtRej_T1;
   IF #s85_StWtPalPresntAtRej THEN #StateNo := 85; END_IF;
END_REGION

REGION Network 35: Actions for STATE Num:85 StWtPalPresntAtRej
   RUNG wire#powerrail
      Contact( #s85_StWtPalPresntAtRej )
      Coil( #qOutput1 )
   END_RUNG
   // the same network as SCL:
   #qOutput1 := #s85_StWtPalPresntAtRej;
END_REGION

REGION Network 36: Transition for STATE Num:90 StWtTTUpStprUp
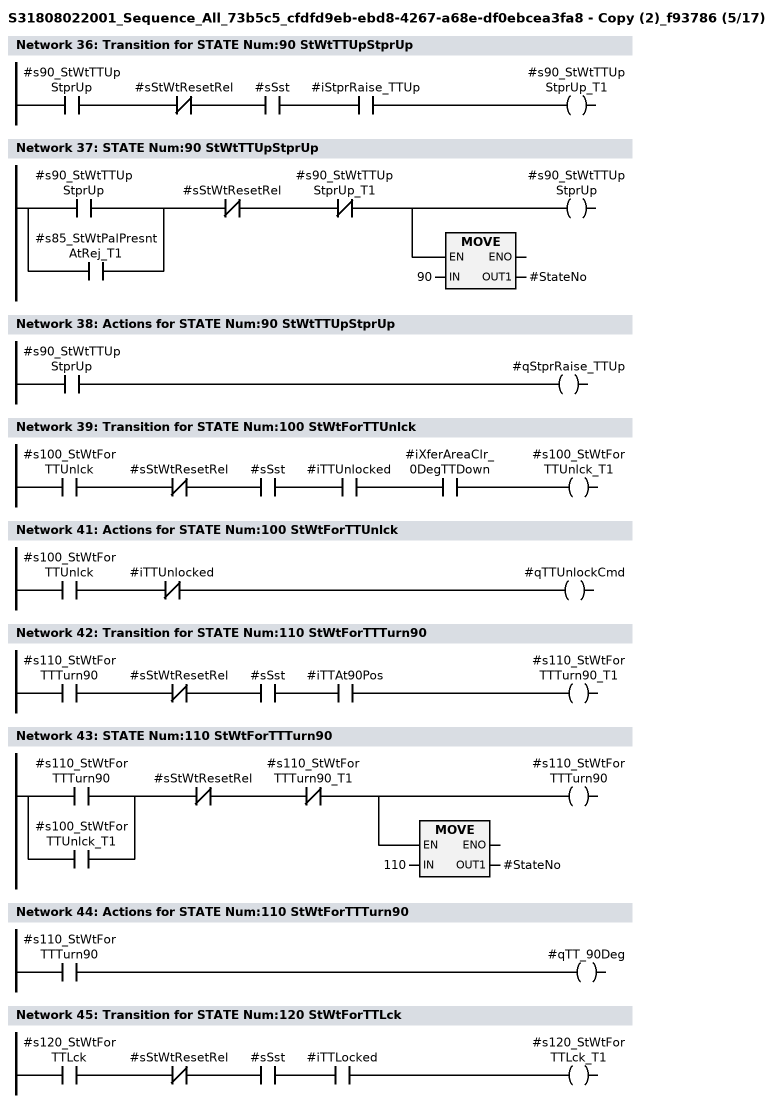
   RUNG wire#powerrail
      Contact( #s90_StWtTTUpStprUp )
      I_Contact( #sStWtResetRel )
      Contact( #sSst )
      Contact( #iStprRaise_TTUp )
      Coil( #s90_StWtTTUpStprUp_T1 )
   END_RUNG
   // the same network as SCL:
   #s90_StWtTTUpStprUp_T1 := #s90_StWtTTUpStprUp AND NOT #sStWtResetRel AND #sSst AND #iStprRaise_TTUp;
END_REGION

REGION Network 37: STATE Num:90 StWtTTUpStprUp
   RUNG wire#powerrail
      Contact( #s90_StWtTTUpStprUp )
      wire#w1
      I_Contact( #sStWtResetRel )
      I_Contact( #s90_StWtTTUpStprUp_T1 )
      wire#w2
      Coil( #s90_StWtTTUpStprUp )
   END_RUNG
   RUNG wire#powerrail
      Contact( #s85_StWtPalPresntAtRej_T1 )
   END_RUNG wire#w1
   RUNG wire#w2
      { S7_GenerateENO := "TRUE" } Move(in := 90, out1 => #StateNo)
   END_RUNG
   // the same network as SCL:
   #s90_StWtTTUpStprUp := (#s90_StWtTTUpStprUp OR #s85_StWtPalPresntAtRej_T1) AND NOT #sStWtResetRel AND NOT #s90_StWtTTUpStprUp_T1;
   IF #s90_StWtTTUpStprUp THEN #StateNo := 90; END_IF;
END_REGION

REGION Network 38: Actions for STATE Num:90 StWtTTUpStprUp
   RUNG wire#powerrail
      Contact( #s90_StWtTTUpStprUp )
      Coil( #qStprRaise_TTUp )
   END_RUNG
   // the same network as SCL:
   #qStprRaise_TTUp := #s90_StWtTTUpStprUp;
END_REGION

REGION Network 39: Transition for STATE Num:100 StWtForTTUnlck
   RUNG wire#powerrail
      Contact( #s100_StWtForTTUnlck )
      I_Contact( #sStWtResetRel )
      Contact( #sSst )
      Contact( #iTTUnlocked )
      Contact( #iXferAreaClr_0DegTTDown )
      Coil( #s100_StWtForTTUnlck_T1 )
   END_RUNG
   // the same network as SCL:
   #s100_StWtForTTUnlck_T1 := #s100_StWtForTTUnlck AND NOT #sStWtResetRel AND #sSst AND #iTTUnlocked AND #iXferAreaClr_0DegTTDown;
END_REGION

NETWORK
TITLE = STATE Num:100 StWtForTTUnlck
      A(;
      O     #s100_StWtForTTUnlck;
      );
      AN    #sStWtResetRel;
      AN    #s100_StWtForTTUnlck_T1;
      =     %L1.0;
      A     %L1.0;
      BLD   102;
      =     #s100_StWtForTTUnlck;
      A     %L1.0;
      JNB   Label_13;
      L     100;
      T     #StateNo;
Label_13:NOP   0;

REGION Network 41: Actions for STATE Num:100 StWtForTTUnlck
   RUNG wire#powerrail
      Contact( #s100_StWtForTTUnlck )
      I_Contact( #iTTUnlocked )
      Coil( #qTTUnlockCmd )
   END_RUNG
   // the same network as SCL:
   #qTTUnlockCmd := #s100_StWtForTTUnlck AND NOT #iTTUnlocked;
END_REGION

REGION Network 42: Transition for STATE Num:110 StWtForTTTurn90
   RUNG wire#powerrail
      Contact( #s110_StWtForTTTurn90 )
      I_Contact( #sStWtResetRel )
      Contact( #sSst )
      Contact( #iTTAt90Pos )
      Coil( #s110_StWtForTTTurn90_T1 )
   END_RUNG
   // the same network as SCL:
   #s110_StWtForTTTurn90_T1 := #s110_StWtForTTTurn90 AND NOT #sStWtResetRel AND #sSst AND #iTTAt90Pos;
END_REGION

REGION Network 43: STATE Num:110 StWtForTTTurn90
   RUNG wire#powerrail
      Contact( #s110_StWtForTTTurn90 )
      wire#w1
      I_Contact( #sStWtResetRel )
      I_Contact( #s110_StWtForTTTurn90_T1 )
      wire#w2
      Coil( #s110_StWtForTTTurn90 )
   END_RUNG
   RUNG wire#powerrail
      Contact( #s100_StWtForTTUnlck_T1 )
   END_RUNG wire#w1
   RUNG wire#w2
      { S7_GenerateENO := "TRUE" } Move(in := 110, out1 => #StateNo)
   END_RUNG
   // the same network as SCL:
   #s110_StWtForTTTurn90 := (#s110_StWtForTTTurn90 OR #s100_StWtForTTUnlck_T1) AND NOT #sStWtResetRel AND NOT #s110_StWtForTTTurn90_T1;
   IF #s110_StWtForTTTurn90 THEN #StateNo := 110; END_IF;
END_REGION

REGION Network 44: Actions for STATE Num:110 StWtForTTTurn90
   RUNG wire#powerrail
      Contact( #s110_StWtForTTTurn90 )
      Coil( #qTT_90Deg )
   END_RUNG
   // the same network as SCL:
   #qTT_90Deg := #s110_StWtForTTTurn90;
END_REGION

REGION Network 45: Transition for STATE Num:120 StWtForTTLck
   RUNG wire#powerrail
      Contact( #s120_StWtForTTLck )
      I_Contact( #sStWtResetRel )
      Contact( #sSst )
      Contact( #iTTLocked )
      Coil( #s120_StWtForTTLck_T1 )
   END_RUNG
   // the same network as SCL:
   #s120_StWtForTTLck_T1 := #s120_StWtForTTLck AND NOT #sStWtResetRel AND #sSst AND #iTTLocked;
END_REGION

REGION Network 46: STATE Num:120 StWtForTTLck
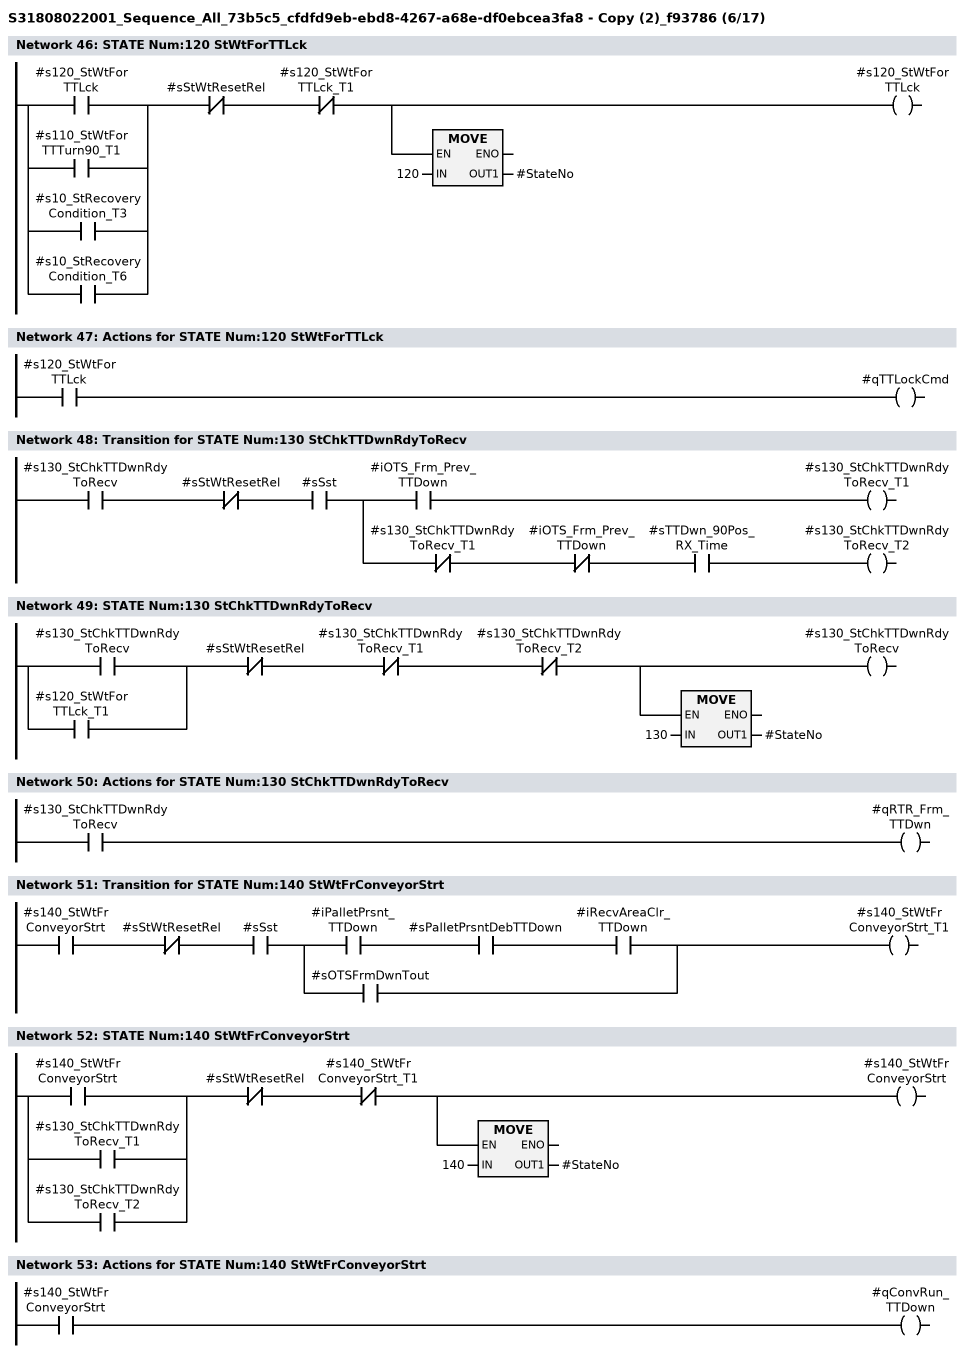
   RUNG wire#powerrail
      Contact( #s120_StWtForTTLck )
      wire#w1
      I_Contact( #sStWtResetRel )
      I_Contact( #s120_StWtForTTLck_T1 )
      wire#w2
      Coil( #s120_StWtForTTLck )
   END_RUNG
   RUNG wire#powerrail
      Contact( #s110_StWtForTTTurn90_T1 )
   END_RUNG wire#w1
   RUNG wire#powerrail
      Contact( #s10_StRecoveryCondition_T3 )
   END_RUNG wire#w1
   RUNG wire#powerrail
      Contact( #s10_StRecoveryCondition_T6 )
   END_RUNG wire#w1
   RUNG wire#w2
      { S7_GenerateENO := "TRUE" } Move(in := 120, out1 => #StateNo)
   END_RUNG
   // the same network as SCL:
   #s120_StWtForTTLck := (#s120_StWtForTTLck OR #s110_StWtForTTTurn90_T1 OR #s10_StRecoveryCondition_T3 OR #s10_StRecoveryCondition_T6) AND NOT #sStWtResetRel AND NOT #s120_StWtForTTLck_T1;
   IF #s120_StWtForTTLck THEN #StateNo := 120; END_IF;
END_REGION

REGION Network 47: Actions for STATE Num:120 StWtForTTLck
   RUNG wire#powerrail
      Contact( #s120_StWtForTTLck )
      Coil( #qTTLockCmd )
   END_RUNG
   // the same network as SCL:
   #qTTLockCmd := #s120_StWtForTTLck;
END_REGION

REGION Network 48: Transition for STATE Num:130 StChkTTDwnRdyToRecv
   RUNG wire#powerrail
      Contact( #s130_StChkTTDwnRdyToRecv )
      I_Contact( #sStWtResetRel )
      Contact( #sSst )
      wire#w1
      Contact( #iOTS_Frm_Prev_TTDown )
      Coil( #s130_StChkTTDwnRdyToRecv_T1 )
   END_RUNG
   RUNG wire#w1
      I_Contact( #s130_StChkTTDwnRdyToRecv_T1 )
      I_Contact( #iOTS_Frm_Prev_TTDown )
      Contact( #sTTDwn_90Pos_RX_Time )
      Coil( #s130_StChkTTDwnRdyToRecv_T2 )
   END_RUNG
   // the same network as SCL:
   #_w1 := #s130_StChkTTDwnRdyToRecv AND NOT #sStWtResetRel AND #sSst;
   #s130_StChkTTDwnRdyToRecv_T1 := #_w1 AND #iOTS_Frm_Prev_TTDown;
   #s130_StChkTTDwnRdyToRecv_T2 := #_w1 AND NOT #s130_StChkTTDwnRdyToRecv_T1 AND NOT #iOTS_Frm_Prev_TTDown AND #sTTDwn_90Pos_RX_Time;
END_REGION

REGION Network 49: STATE Num:130 StChkTTDwnRdyToRecv
   RUNG wire#powerrail
      Contact( #s130_StChkTTDwnRdyToRecv )
      wire#w1
      I_Contact( #sStWtResetRel )
      I_Contact( #s130_StChkTTDwnRdyToRecv_T1 )
      I_Contact( #s130_StChkTTDwnRdyToRecv_T2 )
      wire#w2
      Coil( #s130_StChkTTDwnRdyToRecv )
   END_RUNG
   RUNG wire#powerrail
      Contact( #s120_StWtForTTLck_T1 )
   END_RUNG wire#w1
   RUNG wire#w2
      { S7_GenerateENO := "TRUE" } Move(in := 130, out1 => #StateNo)
   END_RUNG
   // the same network as SCL:
   #s130_StChkTTDwnRdyToRecv := (#s130_StChkTTDwnRdyToRecv OR #s120_StWtForTTLck_T1) AND NOT #sStWtResetRel AND NOT #s130_StChkTTDwnRdyToRecv_T1 AND NOT #s130_StChkTTDwnRdyToRecv_T2;
   IF #s130_StChkTTDwnRdyToRecv THEN #StateNo := 130; END_IF;
END_REGION

REGION Network 50: Actions for STATE Num:130 StChkTTDwnRdyToRecv
   RUNG wire#powerrail
      Contact( #s130_StChkTTDwnRdyToRecv )
      Coil( #qRTR_Frm_TTDwn )
   END_RUNG
   // the same network as SCL:
   #qRTR_Frm_TTDwn := #s130_StChkTTDwnRdyToRecv;
END_REGION

REGION Network 51: Transition for STATE Num:140 StWtFrConveyorStrt
   RUNG wire#powerrail
      Contact( #s140_StWtFrConveyorStrt )
      I_Contact( #sStWtResetRel )
      Contact( #sSst )
      wire#w1
      Contact( #iPalletPrsnt_TTDown )
      Contact( #sPalletPrsntDebTTDown )
      Contact( #iRecvAreaClr_TTDown )
      wire#w2
      Coil( #s140_StWtFrConveyorStrt_T1 )
   END_RUNG
   RUNG wire#w1
      Contact( #sOTSFrmDwnTout )
   END_RUNG wire#w2
   // the same network as SCL:
   #s140_StWtFrConveyorStrt_T1 := #s140_StWtFrConveyorStrt AND NOT #sStWtResetRel AND #sSst AND ((#iPalletPrsnt_TTDown AND #sPalletPrsntDebTTDown AND #iRecvAreaClr_TTDown) OR #sOTSFrmDwnTout);
END_REGION

REGION Network 52: STATE Num:140 StWtFrConveyorStrt
   RUNG wire#powerrail
      Contact( #s140_StWtFrConveyorStrt )
      wire#w1
      I_Contact( #sStWtResetRel )
      I_Contact( #s140_StWtFrConveyorStrt_T1 )
      wire#w2
      Coil( #s140_StWtFrConveyorStrt )
   END_RUNG
   RUNG wire#powerrail
      Contact( #s130_StChkTTDwnRdyToRecv_T1 )
   END_RUNG wire#w1
   RUNG wire#powerrail
      Contact( #s130_StChkTTDwnRdyToRecv_T2 )
   END_RUNG wire#w1
   RUNG wire#w2
      { S7_GenerateENO := "TRUE" } Move(in := 140, out1 => #StateNo)
   END_RUNG
   // the same network as SCL:
   #s140_StWtFrConveyorStrt := (#s140_StWtFrConveyorStrt OR #s130_StChkTTDwnRdyToRecv_T1 OR #s130_StChkTTDwnRdyToRecv_T2) AND NOT #sStWtResetRel AND NOT #s140_StWtFrConveyorStrt_T1;
   IF #s140_StWtFrConveyorStrt THEN #StateNo := 140; END_IF;
END_REGION

REGION Network 53: Actions for STATE Num:140 StWtFrConveyorStrt
   RUNG wire#powerrail
      Contact( #s140_StWtFrConveyorStrt )
      Coil( #qConvRun_TTDown )
   END_RUNG
   // the same network as SCL:
   #qConvRun_TTDown := #s140_StWtFrConveyorStrt;
END_REGION

REGION Network 54: Transition for STATE Num:150 StChkNxtStRdyToRecvTTUp
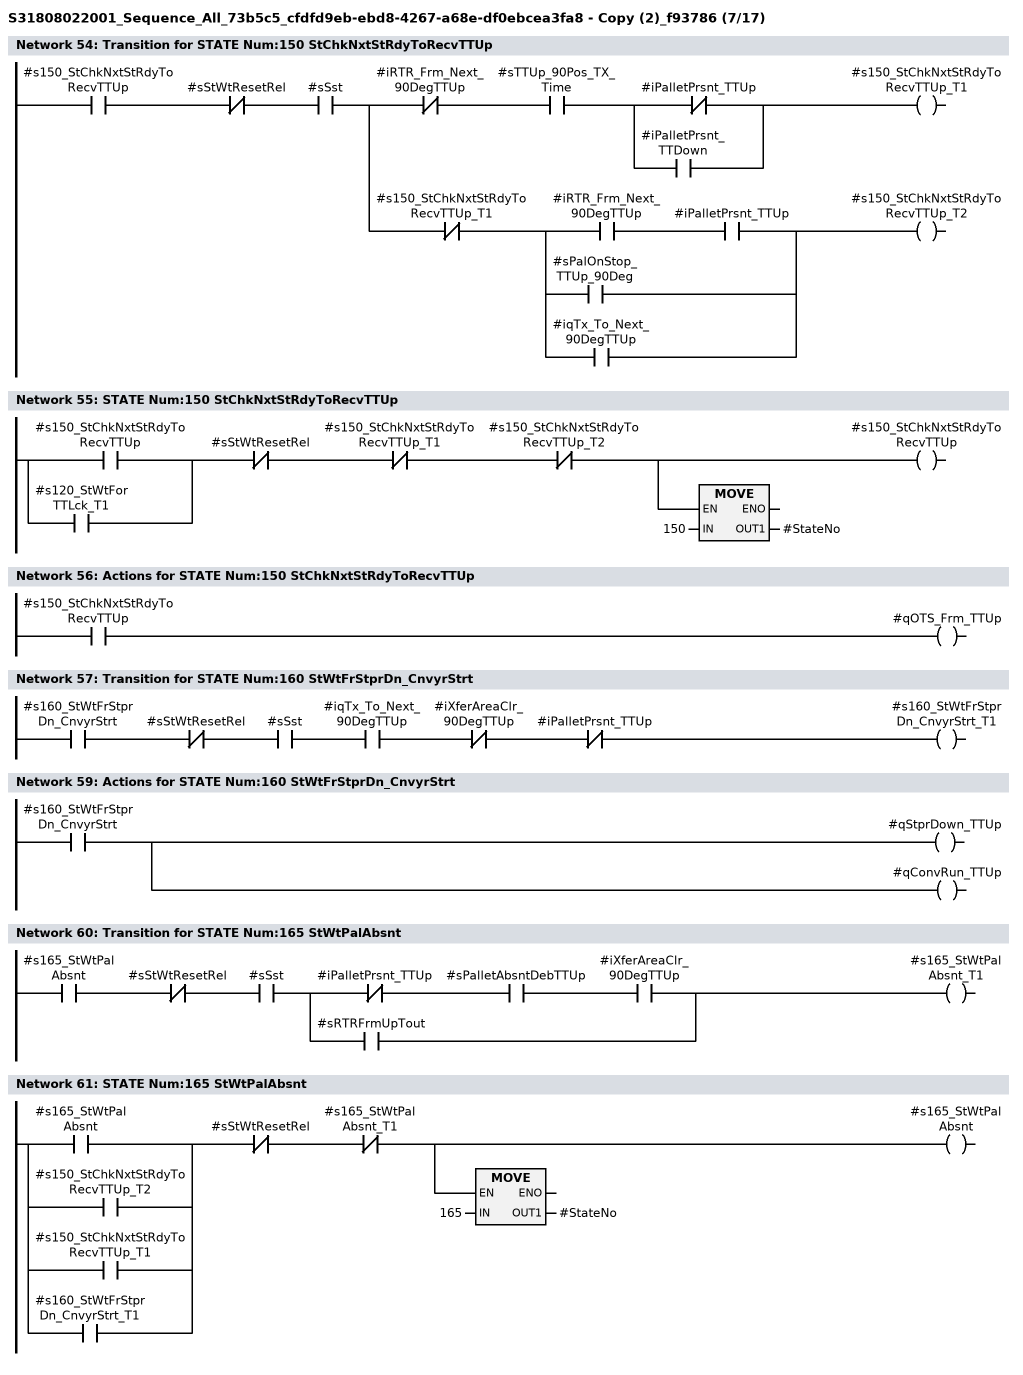
   RUNG wire#powerrail
      Contact( #s150_StChkNxtStRdyToRecvTTUp )
      I_Contact( #sStWtResetRel )
      Contact( #sSst )
      wire#w1
      I_Contact( #iRTR_Frm_Next_90DegTTUp )
      Contact( #sTTUp_90Pos_TX_Time )
      wire#w2
      I_Contact( #iPalletPrsnt_TTUp )
      wire#w3
      Coil( #s150_StChkNxtStRdyToRecvTTUp_T1 )
   END_RUNG
   RUNG wire#w2
      Contact( #iPalletPrsnt_TTDown )
   END_RUNG wire#w3
   RUNG wire#w1
      I_Contact( #s150_StChkNxtStRdyToRecvTTUp_T1 )
      wire#w4
      Contact( #iRTR_Frm_Next_90DegTTUp )
      Contact( #iPalletPrsnt_TTUp )
      wire#w5
      Coil( #s150_StChkNxtStRdyToRecvTTUp_T2 )
   END_RUNG
   RUNG wire#w4
      Contact( #sPalOnStop_TTUp_90Deg )
   END_RUNG wire#w5
   RUNG wire#w4
      Contact( #iqTx_To_Next_90DegTTUp )
   END_RUNG wire#w5
   // the same network as SCL:
   #_w1 := #s150_StChkNxtStRdyToRecvTTUp AND NOT #sStWtResetRel AND #sSst;
   #s150_StChkNxtStRdyToRecvTTUp_T1 := #_w1 AND NOT #iRTR_Frm_Next_90DegTTUp AND #sTTUp_90Pos_TX_Time AND (NOT #iPalletPrsnt_TTUp OR #iPalletPrsnt_TTDown);
   #s150_StChkNxtStRdyToRecvTTUp_T2 := #_w1 AND NOT #s150_StChkNxtStRdyToRecvTTUp_T1 AND ((#iRTR_Frm_Next_90DegTTUp AND #iPalletPrsnt_TTUp) OR #sPalOnStop_TTUp_90Deg OR #iqTx_To_Next_90DegTTUp);
END_REGION

REGION Network 55: STATE Num:150 StChkNxtStRdyToRecvTTUp
   RUNG wire#powerrail
      Contact( #s150_StChkNxtStRdyToRecvTTUp )
      wire#w1
      I_Contact( #sStWtResetRel )
      I_Contact( #s150_StChkNxtStRdyToRecvTTUp_T1 )
      I_Contact( #s150_StChkNxtStRdyToRecvTTUp_T2 )
      wire#w2
      Coil( #s150_StChkNxtStRdyToRecvTTUp )
   END_RUNG
   RUNG wire#powerrail
      Contact( #s120_StWtForTTLck_T1 )
   END_RUNG wire#w1
   RUNG wire#w2
      { S7_GenerateENO := "TRUE" } Move(in := 150, out1 => #StateNo)
   END_RUNG
   // the same network as SCL:
   #s150_StChkNxtStRdyToRecvTTUp := (#s150_StChkNxtStRdyToRecvTTUp OR #s120_StWtForTTLck_T1) AND NOT #sStWtResetRel AND NOT #s150_StChkNxtStRdyToRecvTTUp_T1 AND NOT #s150_StChkNxtStRdyToRecvTTUp_T2;
   IF #s150_StChkNxtStRdyToRecvTTUp THEN #StateNo := 150; END_IF;
END_REGION

REGION Network 56: Actions for STATE Num:150 StChkNxtStRdyToRecvTTUp
   RUNG wire#powerrail
      Contact( #s150_StChkNxtStRdyToRecvTTUp )
      Coil( #qOTS_Frm_TTUp )
   END_RUNG
   // the same network as SCL:
   #qOTS_Frm_TTUp := #s150_StChkNxtStRdyToRecvTTUp;
END_REGION

REGION Network 57: Transition for STATE Num:160 StWtFrStprDn_CnvyrStrt
   RUNG wire#powerrail
      Contact( #s160_StWtFrStprDn_CnvyrStrt )
      I_Contact( #sStWtResetRel )
      Contact( #sSst )
      Contact( #iqTx_To_Next_90DegTTUp )
      I_Contact( #iXferAreaClr_90DegTTUp )
      I_Contact( #iPalletPrsnt_TTUp )
      Coil( #s160_StWtFrStprDn_CnvyrStrt_T1 )
   END_RUNG
   // the same network as SCL:
   #s160_StWtFrStprDn_CnvyrStrt_T1 := #s160_StWtFrStprDn_CnvyrStrt AND NOT #sStWtResetRel AND #sSst AND #iqTx_To_Next_90DegTTUp AND NOT #iXferAreaClr_90DegTTUp AND NOT #iPalletPrsnt_TTUp;
END_REGION

NETWORK
TITLE = STATE Num:160 StWtFrStprDn_CnvyrStrt
      A(;
      O     #s160_StWtFrStprDn_CnvyrStrt;
//wrong transition variable removed
      );
      AN    #sStWtResetRel;
      AN    #s160_StWtFrStprDn_CnvyrStrt_T1;
      =     %L1.0;
      A     %L1.0;
      BLD   102;
      =     #s160_StWtFrStprDn_CnvyrStrt;
      A     %L1.0;
      JNB   Label_19;
      L     160;
      T     #StateNo;
Label_19:NOP   0;

REGION Network 59: Actions for STATE Num:160 StWtFrStprDn_CnvyrStrt
   RUNG wire#powerrail
      Contact( #s160_StWtFrStprDn_CnvyrStrt )
      wire#w1
      Coil( #qStprDown_TTUp )
   END_RUNG
   RUNG wire#w1
      Coil( #qConvRun_TTUp )
   END_RUNG
   // the same network as SCL:
   #qStprDown_TTUp := #s160_StWtFrStprDn_CnvyrStrt;
   #qConvRun_TTUp := #s160_StWtFrStprDn_CnvyrStrt;
END_REGION

REGION Network 60: Transition for STATE Num:165 StWtPalAbsnt
   RUNG wire#powerrail
      Contact( #s165_StWtPalAbsnt )
      I_Contact( #sStWtResetRel )
      Contact( #sSst )
      wire#w1
      I_Contact( #iPalletPrsnt_TTUp )
      Contact( #sPalletAbsntDebTTUp )
      Contact( #iXferAreaClr_90DegTTUp )
      wire#w2
      Coil( #s165_StWtPalAbsnt_T1 )
   END_RUNG
   RUNG wire#w1
      Contact( #sRTRFrmUpTout )
   END_RUNG wire#w2
   // the same network as SCL:
   #s165_StWtPalAbsnt_T1 := #s165_StWtPalAbsnt AND NOT #sStWtResetRel AND #sSst AND ((NOT #iPalletPrsnt_TTUp AND #sPalletAbsntDebTTUp AND #iXferAreaClr_90DegTTUp) OR #sRTRFrmUpTout);
END_REGION

REGION Network 61: STATE Num:165 StWtPalAbsnt
   RUNG wire#powerrail
      Contact( #s165_StWtPalAbsnt )
      wire#w1
      I_Contact( #sStWtResetRel )
      I_Contact( #s165_StWtPalAbsnt_T1 )
      wire#w2
      Coil( #s165_StWtPalAbsnt )
   END_RUNG
   RUNG wire#powerrail
      Contact( #s150_StChkNxtStRdyToRecvTTUp_T2 )
   END_RUNG wire#w1
   RUNG wire#powerrail
      Contact( #s150_StChkNxtStRdyToRecvTTUp_T1 )
   END_RUNG wire#w1
   RUNG wire#powerrail
      Contact( #s160_StWtFrStprDn_CnvyrStrt_T1 )
   END_RUNG wire#w1
   RUNG wire#w2
      { S7_GenerateENO := "TRUE" } Move(in := 165, out1 => #StateNo)
   END_RUNG
   // the same network as SCL:
   #s165_StWtPalAbsnt := (#s165_StWtPalAbsnt OR #s150_StChkNxtStRdyToRecvTTUp_T2 OR #s150_StChkNxtStRdyToRecvTTUp_T1 OR #s160_StWtFrStprDn_CnvyrStrt_T1) AND NOT #sStWtResetRel AND NOT #s165_StWtPalAbsnt_T1;
   IF #s165_StWtPalAbsnt THEN #StateNo := 165; END_IF;
END_REGION

REGION Network 62: Actions for STATE Num:165 StWtPalAbsnt
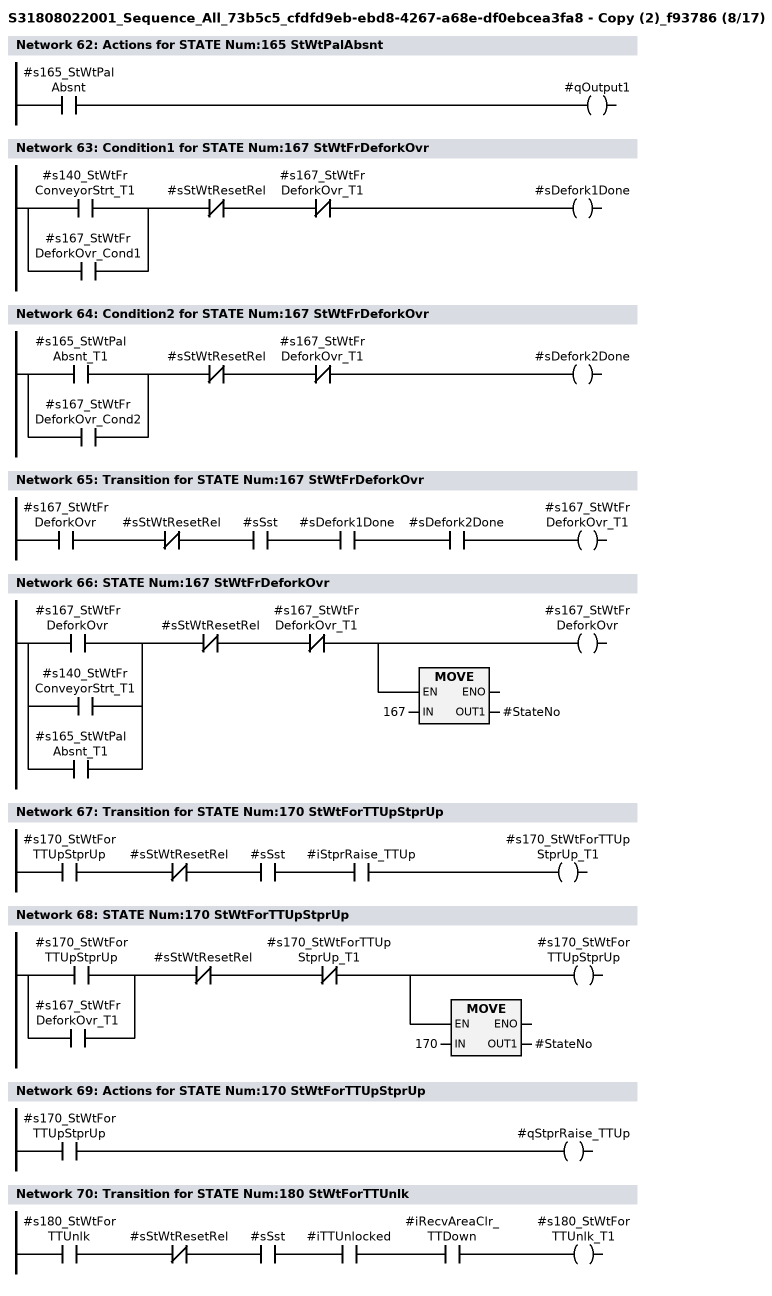
   RUNG wire#powerrail
      Contact( #s165_StWtPalAbsnt )
      Coil( #qOutput1 )
   END_RUNG
   // the same network as SCL:
   #qOutput1 := #s165_StWtPalAbsnt;
END_REGION

REGION Network 63: Condition1 for STATE Num:167 StWtFrDeforkOvr
   RUNG wire#powerrail
      Contact( #s140_StWtFrConveyorStrt_T1 )
      wire#w1
      I_Contact( #sStWtResetRel )
      I_Contact( #s167_StWtFrDeforkOvr_T1 )
      Coil( #sDefork1Done )
   END_RUNG
   RUNG wire#powerrail
      Contact( #s167_StWtFrDeforkOvr_Cond1 )
   END_RUNG wire#w1
   // the same network as SCL:
   #sDefork1Done := (#s140_StWtFrConveyorStrt_T1 OR #s167_StWtFrDeforkOvr_Cond1) AND NOT #sStWtResetRel AND NOT #s167_StWtFrDeforkOvr_T1;
END_REGION

REGION Network 64: Condition2 for STATE Num:167 StWtFrDeforkOvr
   RUNG wire#powerrail
      Contact( #s165_StWtPalAbsnt_T1 )
      wire#w1
      I_Contact( #sStWtResetRel )
      I_Contact( #s167_StWtFrDeforkOvr_T1 )
      Coil( #sDefork2Done )
   END_RUNG
   RUNG wire#powerrail
      Contact( #s167_StWtFrDeforkOvr_Cond2 )
   END_RUNG wire#w1
   // the same network as SCL:
   #sDefork2Done := (#s165_StWtPalAbsnt_T1 OR #s167_StWtFrDeforkOvr_Cond2) AND NOT #sStWtResetRel AND NOT #s167_StWtFrDeforkOvr_T1;
END_REGION

REGION Network 65: Transition for STATE Num:167 StWtFrDeforkOvr
   RUNG wire#powerrail
      Contact( #s167_StWtFrDeforkOvr )
      I_Contact( #sStWtResetRel )
      Contact( #sSst )
      Contact( #sDefork1Done )
      Contact( #sDefork2Done )
      Coil( #s167_StWtFrDeforkOvr_T1 )
   END_RUNG
   // the same network as SCL:
   #s167_StWtFrDeforkOvr_T1 := #s167_StWtFrDeforkOvr AND NOT #sStWtResetRel AND #sSst AND #sDefork1Done AND #sDefork2Done;
END_REGION

REGION Network 66: STATE Num:167 StWtFrDeforkOvr
   RUNG wire#powerrail
      Contact( #s167_StWtFrDeforkOvr )
      wire#w1
      I_Contact( #sStWtResetRel )
      I_Contact( #s167_StWtFrDeforkOvr_T1 )
      wire#w2
      Coil( #s167_StWtFrDeforkOvr )
   END_RUNG
   RUNG wire#powerrail
      Contact( #s140_StWtFrConveyorStrt_T1 )
   END_RUNG wire#w1
   RUNG wire#powerrail
      Contact( #s165_StWtPalAbsnt_T1 )
   END_RUNG wire#w1
   RUNG wire#w2
      { S7_GenerateENO := "TRUE" } Move(in := 167, out1 => #StateNo)
   END_RUNG
   // the same network as SCL:
   #s167_StWtFrDeforkOvr := (#s167_StWtFrDeforkOvr OR #s140_StWtFrConveyorStrt_T1 OR #s165_StWtPalAbsnt_T1) AND NOT #sStWtResetRel AND NOT #s167_StWtFrDeforkOvr_T1;
   IF #s167_StWtFrDeforkOvr THEN #StateNo := 167; END_IF;
END_REGION

REGION Network 67: Transition for STATE Num:170 StWtForTTUpStprUp
   RUNG wire#powerrail
      Contact( #s170_StWtForTTUpStprUp )
      I_Contact( #sStWtResetRel )
      Contact( #sSst )
      Contact( #iStprRaise_TTUp )
      Coil( #s170_StWtForTTUpStprUp_T1 )
   END_RUNG
   // the same network as SCL:
   #s170_StWtForTTUpStprUp_T1 := #s170_StWtForTTUpStprUp AND NOT #sStWtResetRel AND #sSst AND #iStprRaise_TTUp;
END_REGION

REGION Network 68: STATE Num:170 StWtForTTUpStprUp
   RUNG wire#powerrail
      Contact( #s170_StWtForTTUpStprUp )
      wire#w1
      I_Contact( #sStWtResetRel )
      I_Contact( #s170_StWtForTTUpStprUp_T1 )
      wire#w2
      Coil( #s170_StWtForTTUpStprUp )
   END_RUNG
   RUNG wire#powerrail
      Contact( #s167_StWtFrDeforkOvr_T1 )
   END_RUNG wire#w1
   RUNG wire#w2
      { S7_GenerateENO := "TRUE" } Move(in := 170, out1 => #StateNo)
   END_RUNG
   // the same network as SCL:
   #s170_StWtForTTUpStprUp := (#s170_StWtForTTUpStprUp OR #s167_StWtFrDeforkOvr_T1) AND NOT #sStWtResetRel AND NOT #s170_StWtForTTUpStprUp_T1;
   IF #s170_StWtForTTUpStprUp THEN #StateNo := 170; END_IF;
END_REGION

REGION Network 69: Actions for STATE Num:170 StWtForTTUpStprUp
   RUNG wire#powerrail
      Contact( #s170_StWtForTTUpStprUp )
      Coil( #qStprRaise_TTUp )
   END_RUNG
   // the same network as SCL:
   #qStprRaise_TTUp := #s170_StWtForTTUpStprUp;
END_REGION

REGION Network 70: Transition for STATE Num:180 StWtForTTUnlk
   RUNG wire#powerrail
      Contact( #s180_StWtForTTUnlk )
      I_Contact( #sStWtResetRel )
      Contact( #sSst )
      Contact( #iTTUnlocked )
      Contact( #iRecvAreaClr_TTDown )
      Coil( #s180_StWtForTTUnlk_T1 )
   END_RUNG
   // the same network as SCL:
   #s180_StWtForTTUnlk_T1 := #s180_StWtForTTUnlk AND NOT #sStWtResetRel AND #sSst AND #iTTUnlocked AND #iRecvAreaClr_TTDown;
END_REGION

REGION Network 71: STATE Num:180 StWtForTTUnlk
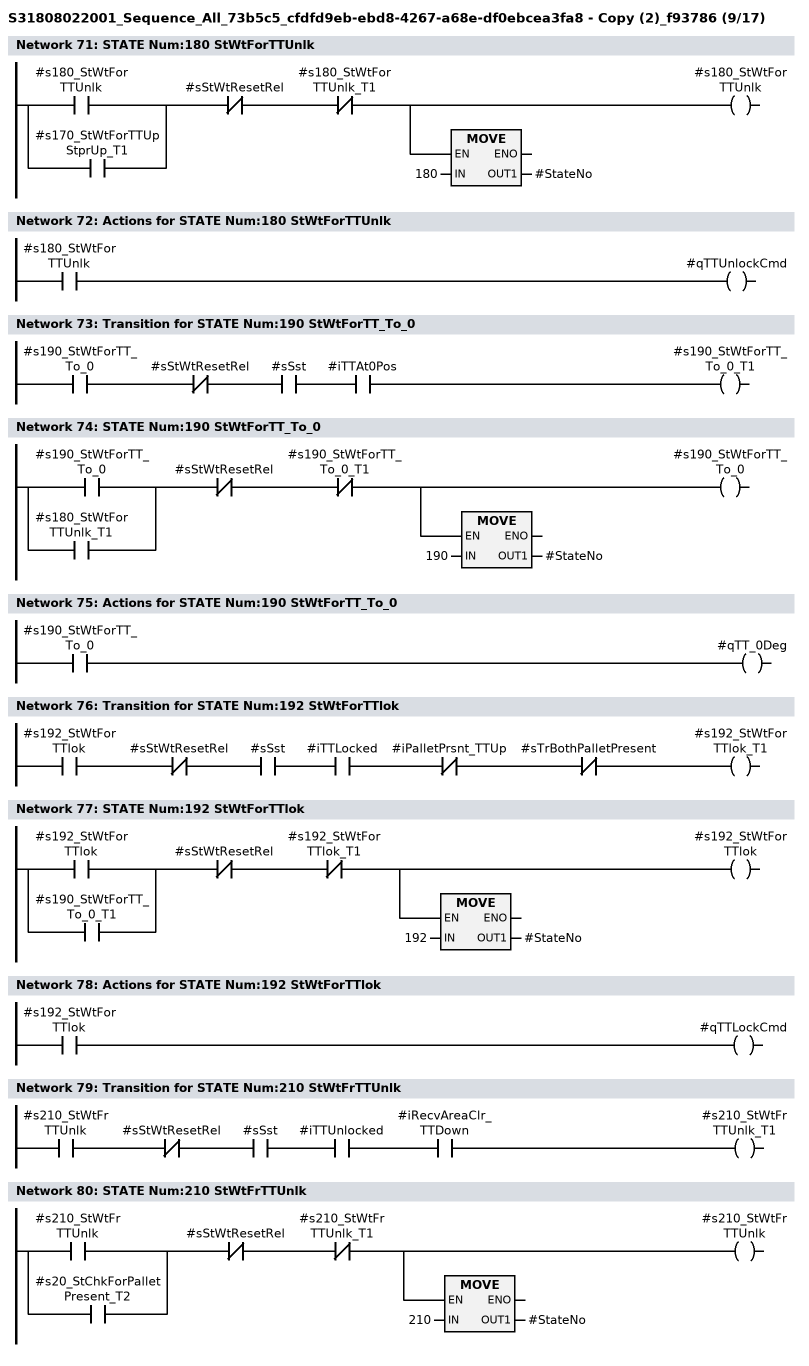
   RUNG wire#powerrail
      Contact( #s180_StWtForTTUnlk )
      wire#w1
      I_Contact( #sStWtResetRel )
      I_Contact( #s180_StWtForTTUnlk_T1 )
      wire#w2
      Coil( #s180_StWtForTTUnlk )
   END_RUNG
   RUNG wire#powerrail
      Contact( #s170_StWtForTTUpStprUp_T1 )
   END_RUNG wire#w1
   RUNG wire#w2
      { S7_GenerateENO := "TRUE" } Move(in := 180, out1 => #StateNo)
   END_RUNG
   // the same network as SCL:
   #s180_StWtForTTUnlk := (#s180_StWtForTTUnlk OR #s170_StWtForTTUpStprUp_T1) AND NOT #sStWtResetRel AND NOT #s180_StWtForTTUnlk_T1;
   IF #s180_StWtForTTUnlk THEN #StateNo := 180; END_IF;
END_REGION

REGION Network 72: Actions for STATE Num:180 StWtForTTUnlk
   RUNG wire#powerrail
      Contact( #s180_StWtForTTUnlk )
      Coil( #qTTUnlockCmd )
   END_RUNG
   // the same network as SCL:
   #qTTUnlockCmd := #s180_StWtForTTUnlk;
END_REGION

REGION Network 73: Transition for STATE Num:190 StWtForTT_To_0
   RUNG wire#powerrail
      Contact( #s190_StWtForTT_To_0 )
      I_Contact( #sStWtResetRel )
      Contact( #sSst )
      Contact( #iTTAt0Pos )
      Coil( #s190_StWtForTT_To_0_T1 )
   END_RUNG
   // the same network as SCL:
   #s190_StWtForTT_To_0_T1 := #s190_StWtForTT_To_0 AND NOT #sStWtResetRel AND #sSst AND #iTTAt0Pos;
END_REGION

REGION Network 74: STATE Num:190 StWtForTT_To_0
   RUNG wire#powerrail
      Contact( #s190_StWtForTT_To_0 )
      wire#w1
      I_Contact( #sStWtResetRel )
      I_Contact( #s190_StWtForTT_To_0_T1 )
      wire#w2
      Coil( #s190_StWtForTT_To_0 )
   END_RUNG
   RUNG wire#powerrail
      Contact( #s180_StWtForTTUnlk_T1 )
   END_RUNG wire#w1
   RUNG wire#w2
      { S7_GenerateENO := "TRUE" } Move(in := 190, out1 => #StateNo)
   END_RUNG
   // the same network as SCL:
   #s190_StWtForTT_To_0 := (#s190_StWtForTT_To_0 OR #s180_StWtForTTUnlk_T1) AND NOT #sStWtResetRel AND NOT #s190_StWtForTT_To_0_T1;
   IF #s190_StWtForTT_To_0 THEN #StateNo := 190; END_IF;
END_REGION

REGION Network 75: Actions for STATE Num:190 StWtForTT_To_0
   RUNG wire#powerrail
      Contact( #s190_StWtForTT_To_0 )
      Coil( #qTT_0Deg )
   END_RUNG
   // the same network as SCL:
   #qTT_0Deg := #s190_StWtForTT_To_0;
END_REGION

REGION Network 76: Transition for STATE Num:192 StWtForTTlok
   RUNG wire#powerrail
      Contact( #s192_StWtForTTlok )
      I_Contact( #sStWtResetRel )
      Contact( #sSst )
      Contact( #iTTLocked )
      I_Contact( #iPalletPrsnt_TTUp )
      I_Contact( #sTrBothPalletPresent )
      Coil( #s192_StWtForTTlok_T1 )
   END_RUNG
   // the same network as SCL:
   #s192_StWtForTTlok_T1 := #s192_StWtForTTlok AND NOT #sStWtResetRel AND #sSst AND #iTTLocked AND NOT #iPalletPrsnt_TTUp AND NOT #sTrBothPalletPresent;
END_REGION

REGION Network 77: STATE Num:192 StWtForTTlok
   RUNG wire#powerrail
      Contact( #s192_StWtForTTlok )
      wire#w1
      I_Contact( #sStWtResetRel )
      I_Contact( #s192_StWtForTTlok_T1 )
      wire#w2
      Coil( #s192_StWtForTTlok )
   END_RUNG
   RUNG wire#powerrail
      Contact( #s190_StWtForTT_To_0_T1 )
   END_RUNG wire#w1
   RUNG wire#w2
      { S7_GenerateENO := "TRUE" } Move(in := 192, out1 => #StateNo)
   END_RUNG
   // the same network as SCL:
   #s192_StWtForTTlok := (#s192_StWtForTTlok OR #s190_StWtForTT_To_0_T1) AND NOT #sStWtResetRel AND NOT #s192_StWtForTTlok_T1;
   IF #s192_StWtForTTlok THEN #StateNo := 192; END_IF;
END_REGION

REGION Network 78: Actions for STATE Num:192 StWtForTTlok
   RUNG wire#powerrail
      Contact( #s192_StWtForTTlok )
      Coil( #qTTLockCmd )
   END_RUNG
   // the same network as SCL:
   #qTTLockCmd := #s192_StWtForTTlok;
END_REGION

REGION Network 79: Transition for STATE Num:210 StWtFrTTUnlk
   RUNG wire#powerrail
      Contact( #s210_StWtFrTTUnlk )
      I_Contact( #sStWtResetRel )
      Contact( #sSst )
      Contact( #iTTUnlocked )
      Contact( #iRecvAreaClr_TTDown )
      Coil( #s210_StWtFrTTUnlk_T1 )
   END_RUNG
   // the same network as SCL:
   #s210_StWtFrTTUnlk_T1 := #s210_StWtFrTTUnlk AND NOT #sStWtResetRel AND #sSst AND #iTTUnlocked AND #iRecvAreaClr_TTDown;
END_REGION

REGION Network 80: STATE Num:210 StWtFrTTUnlk
   RUNG wire#powerrail
      Contact( #s210_StWtFrTTUnlk )
      wire#w1
      I_Contact( #sStWtResetRel )
      I_Contact( #s210_StWtFrTTUnlk_T1 )
      wire#w2
      Coil( #s210_StWtFrTTUnlk )
   END_RUNG
   RUNG wire#powerrail
      Contact( #s20_StChkForPalletPresent_T2 )
   END_RUNG wire#w1
   RUNG wire#w2
      { S7_GenerateENO := "TRUE" } Move(in := 210, out1 => #StateNo)
   END_RUNG
   // the same network as SCL:
   #s210_StWtFrTTUnlk := (#s210_StWtFrTTUnlk OR #s20_StChkForPalletPresent_T2) AND NOT #sStWtResetRel AND NOT #s210_StWtFrTTUnlk_T1;
   IF #s210_StWtFrTTUnlk THEN #StateNo := 210; END_IF;
END_REGION

REGION Network 81: Actions for STATE Num:210 StWtFrTTUnlk
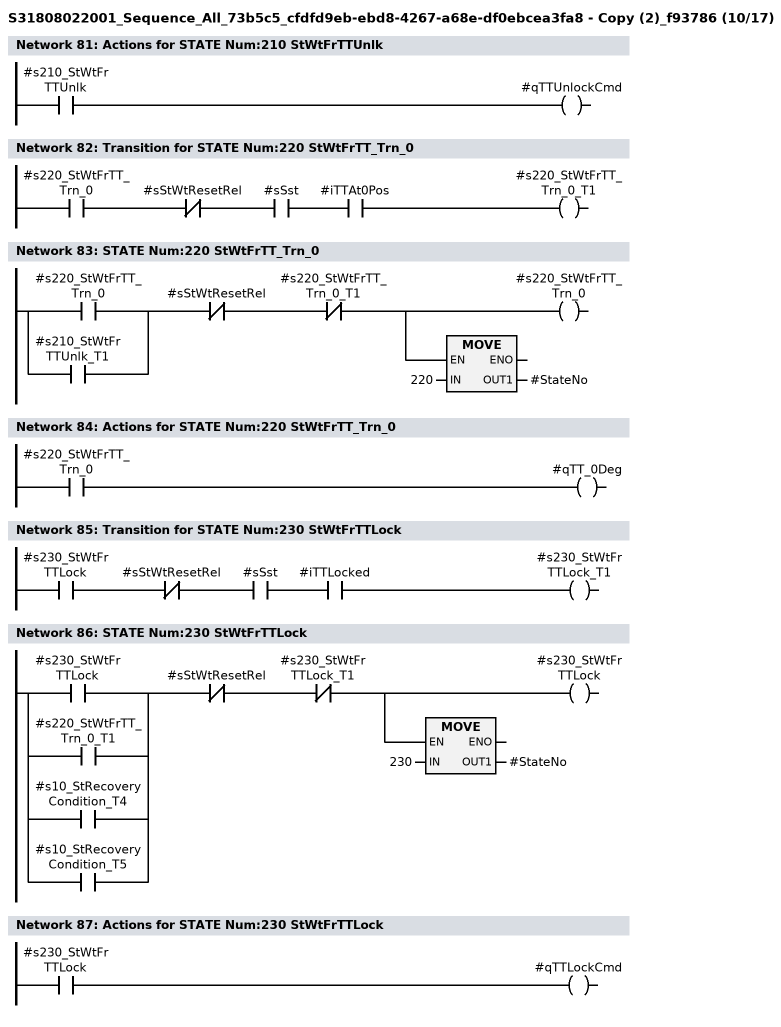
   RUNG wire#powerrail
      Contact( #s210_StWtFrTTUnlk )
      Coil( #qTTUnlockCmd )
   END_RUNG
   // the same network as SCL:
   #qTTUnlockCmd := #s210_StWtFrTTUnlk;
END_REGION

REGION Network 82: Transition for STATE Num:220 StWtFrTT_Trn_0
   RUNG wire#powerrail
      Contact( #s220_StWtFrTT_Trn_0 )
      I_Contact( #sStWtResetRel )
      Contact( #sSst )
      Contact( #iTTAt0Pos )
      Coil( #s220_StWtFrTT_Trn_0_T1 )
   END_RUNG
   // the same network as SCL:
   #s220_StWtFrTT_Trn_0_T1 := #s220_StWtFrTT_Trn_0 AND NOT #sStWtResetRel AND #sSst AND #iTTAt0Pos;
END_REGION

REGION Network 83: STATE Num:220 StWtFrTT_Trn_0
   RUNG wire#powerrail
      Contact( #s220_StWtFrTT_Trn_0 )
      wire#w1
      I_Contact( #sStWtResetRel )
      I_Contact( #s220_StWtFrTT_Trn_0_T1 )
      wire#w2
      Coil( #s220_StWtFrTT_Trn_0 )
   END_RUNG
   RUNG wire#powerrail
      Contact( #s210_StWtFrTTUnlk_T1 )
   END_RUNG wire#w1
   RUNG wire#w2
      { S7_GenerateENO := "TRUE" } Move(in := 220, out1 => #StateNo)
   END_RUNG
   // the same network as SCL:
   #s220_StWtFrTT_Trn_0 := (#s220_StWtFrTT_Trn_0 OR #s210_StWtFrTTUnlk_T1) AND NOT #sStWtResetRel AND NOT #s220_StWtFrTT_Trn_0_T1;
   IF #s220_StWtFrTT_Trn_0 THEN #StateNo := 220; END_IF;
END_REGION

REGION Network 84: Actions for STATE Num:220 StWtFrTT_Trn_0
   RUNG wire#powerrail
      Contact( #s220_StWtFrTT_Trn_0 )
      Coil( #qTT_0Deg )
   END_RUNG
   // the same network as SCL:
   #qTT_0Deg := #s220_StWtFrTT_Trn_0;
END_REGION

REGION Network 85: Transition for STATE Num:230 StWtFrTTLock
   RUNG wire#powerrail
      Contact( #s230_StWtFrTTLock )
      I_Contact( #sStWtResetRel )
      Contact( #sSst )
      Contact( #iTTLocked )
      Coil( #s230_StWtFrTTLock_T1 )
   END_RUNG
   // the same network as SCL:
   #s230_StWtFrTTLock_T1 := #s230_StWtFrTTLock AND NOT #sStWtResetRel AND #sSst AND #iTTLocked;
END_REGION

REGION Network 86: STATE Num:230 StWtFrTTLock
   RUNG wire#powerrail
      Contact( #s230_StWtFrTTLock )
      wire#w1
      I_Contact( #sStWtResetRel )
      I_Contact( #s230_StWtFrTTLock_T1 )
      wire#w2
      Coil( #s230_StWtFrTTLock )
   END_RUNG
   RUNG wire#powerrail
      Contact( #s220_StWtFrTT_Trn_0_T1 )
   END_RUNG wire#w1
   RUNG wire#powerrail
      Contact( #s10_StRecoveryCondition_T4 )
   END_RUNG wire#w1
   RUNG wire#powerrail
      Contact( #s10_StRecoveryCondition_T5 )
   END_RUNG wire#w1
   RUNG wire#w2
      { S7_GenerateENO := "TRUE" } Move(in := 230, out1 => #StateNo)
   END_RUNG
   // the same network as SCL:
   #s230_StWtFrTTLock := (#s230_StWtFrTTLock OR #s220_StWtFrTT_Trn_0_T1 OR #s10_StRecoveryCondition_T4 OR #s10_StRecoveryCondition_T5) AND NOT #sStWtResetRel AND NOT #s230_StWtFrTTLock_T1;
   IF #s230_StWtFrTTLock THEN #StateNo := 230; END_IF;
END_REGION

REGION Network 87: Actions for STATE Num:230 StWtFrTTLock
   RUNG wire#powerrail
      Contact( #s230_StWtFrTTLock )
      Coil( #qTTLockCmd )
   END_RUNG
   // the same network as SCL:
   #qTTLockCmd := #s230_StWtFrTTLock;
END_REGION

REGION Network 88: Transition for STATE Num:240 StWtFRTRNxtStnTTDown
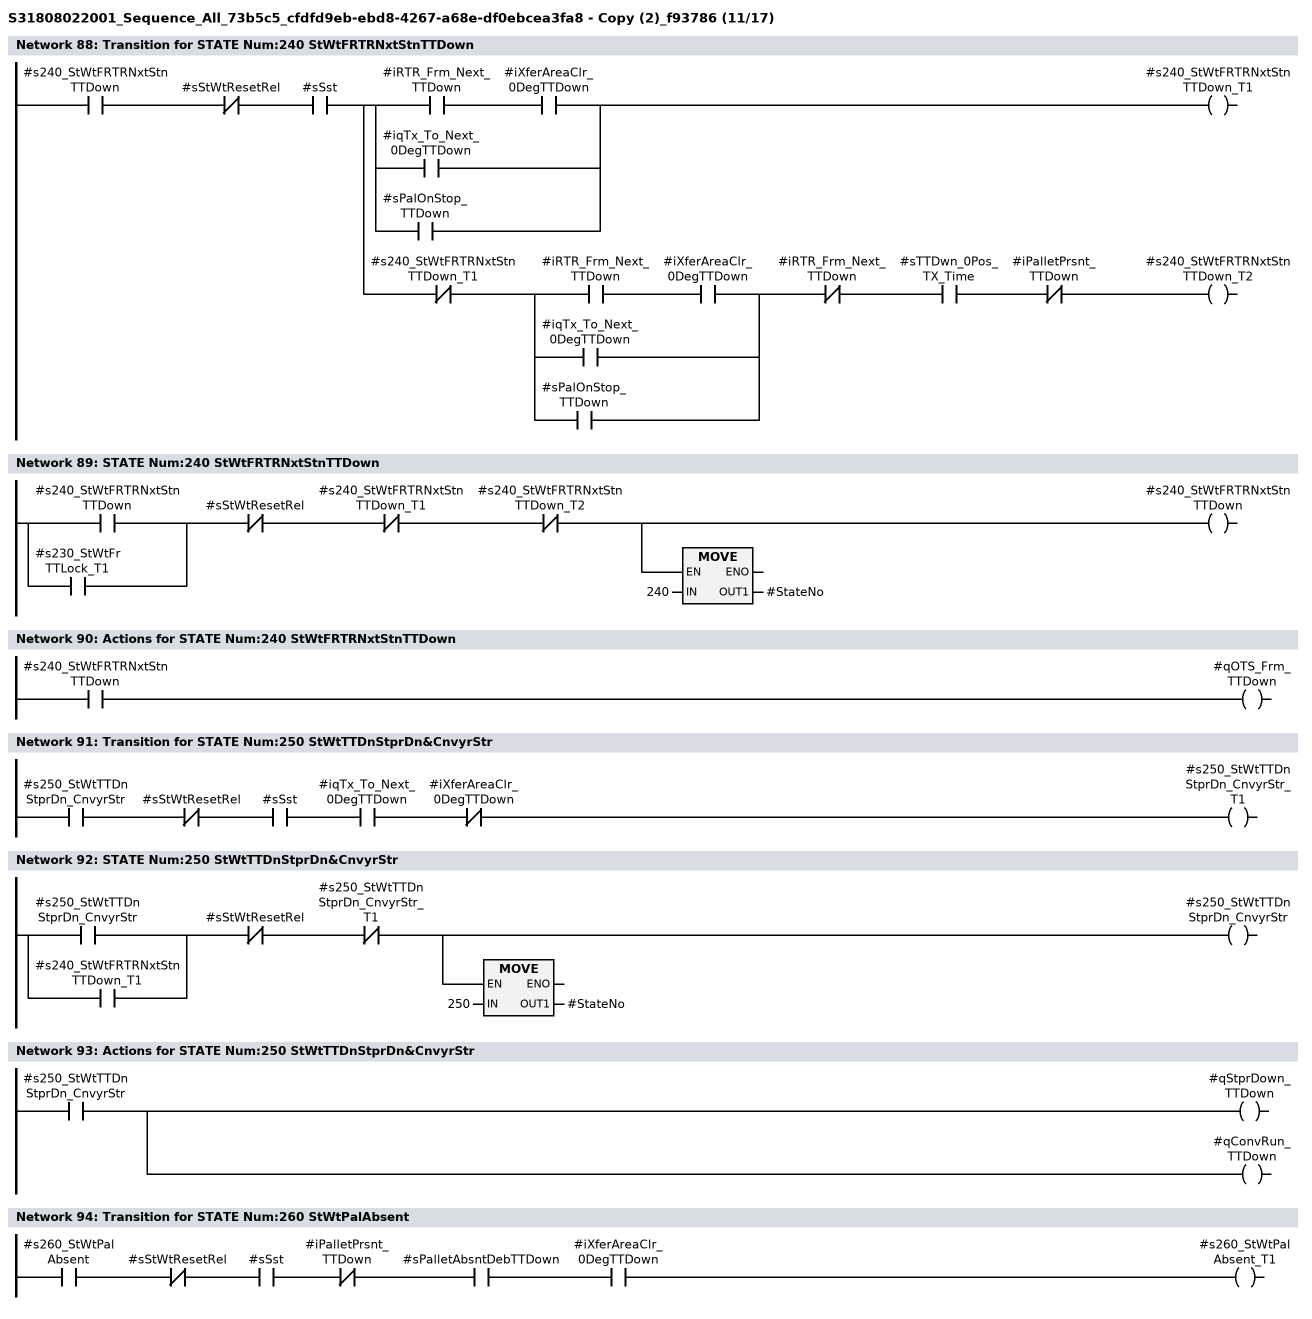
   RUNG wire#powerrail
      Contact( #s240_StWtFRTRNxtStnTTDown )
      I_Contact( #sStWtResetRel )
      Contact( #sSst )
      wire#w1
      Contact( #iRTR_Frm_Next_TTDown )
      Contact( #iXferAreaClr_0DegTTDown )
      wire#w2
      Coil( #s240_StWtFRTRNxtStnTTDown_T1 )
   END_RUNG
   RUNG wire#w1
      Contact( #iqTx_To_Next_0DegTTDown )
   END_RUNG wire#w2
   RUNG wire#w1
      Contact( #sPalOnStop_TTDown )
   END_RUNG wire#w2
   RUNG wire#w1
      I_Contact( #s240_StWtFRTRNxtStnTTDown_T1 )
      wire#w3
      Contact( #iRTR_Frm_Next_TTDown )
      Contact( #iXferAreaClr_0DegTTDown )
      wire#w4
      I_Contact( #iRTR_Frm_Next_TTDown )
      Contact( #sTTDwn_0Pos_TX_Time )
      I_Contact( #iPalletPrsnt_TTDown )
      Coil( #s240_StWtFRTRNxtStnTTDown_T2 )
   END_RUNG
   RUNG wire#w3
      Contact( #iqTx_To_Next_0DegTTDown )
   END_RUNG wire#w4
   RUNG wire#w3
      Contact( #sPalOnStop_TTDown )
   END_RUNG wire#w4
   // the same network as SCL:
   #_w1 := #s240_StWtFRTRNxtStnTTDown AND NOT #sStWtResetRel AND #sSst;
   #s240_StWtFRTRNxtStnTTDown_T1 := #_w1 AND ((#iRTR_Frm_Next_TTDown AND #iXferAreaClr_0DegTTDown) OR #iqTx_To_Next_0DegTTDown OR #sPalOnStop_TTDown);
   #s240_StWtFRTRNxtStnTTDown_T2 := #_w1 AND NOT #s240_StWtFRTRNxtStnTTDown_T1 AND ((#iRTR_Frm_Next_TTDown AND #iXferAreaClr_0DegTTDown) OR #iqTx_To_Next_0DegTTDown OR #sPalOnStop_TTDown) AND NOT #iRTR_Frm_Next_TTDown AND #sTTDwn_0Pos_TX_Time AND NOT #iPalletPrsnt_TTDown;
END_REGION

REGION Network 89: STATE Num:240 StWtFRTRNxtStnTTDown
   RUNG wire#powerrail
      Contact( #s240_StWtFRTRNxtStnTTDown )
      wire#w1
      I_Contact( #sStWtResetRel )
      I_Contact( #s240_StWtFRTRNxtStnTTDown_T1 )
      I_Contact( #s240_StWtFRTRNxtStnTTDown_T2 )
      wire#w2
      Coil( #s240_StWtFRTRNxtStnTTDown )
   END_RUNG
   RUNG wire#powerrail
      Contact( #s230_StWtFrTTLock_T1 )
   END_RUNG wire#w1
   RUNG wire#w2
      { S7_GenerateENO := "TRUE" } Move(in := 240, out1 => #StateNo)
   END_RUNG
   // the same network as SCL:
   #s240_StWtFRTRNxtStnTTDown := (#s240_StWtFRTRNxtStnTTDown OR #s230_StWtFrTTLock_T1) AND NOT #sStWtResetRel AND NOT #s240_StWtFRTRNxtStnTTDown_T1 AND NOT #s240_StWtFRTRNxtStnTTDown_T2;
   IF #s240_StWtFRTRNxtStnTTDown THEN #StateNo := 240; END_IF;
END_REGION

REGION Network 90: Actions for STATE Num:240 StWtFRTRNxtStnTTDown
   RUNG wire#powerrail
      Contact( #s240_StWtFRTRNxtStnTTDown )
      Coil( #qOTS_Frm_TTDown )
   END_RUNG
   // the same network as SCL:
   #qOTS_Frm_TTDown := #s240_StWtFRTRNxtStnTTDown;
END_REGION

REGION Network 91: Transition for STATE Num:250 StWtTTDnStprDn&CnvyrStr
   RUNG wire#powerrail
      Contact( #s250_StWtTTDnStprDn_CnvyrStr )
      I_Contact( #sStWtResetRel )
      Contact( #sSst )
      Contact( #iqTx_To_Next_0DegTTDown )
      I_Contact( #iXferAreaClr_0DegTTDown )
      Coil( #s250_StWtTTDnStprDn_CnvyrStr_T1 )
   END_RUNG
   // the same network as SCL:
   #s250_StWtTTDnStprDn_CnvyrStr_T1 := #s250_StWtTTDnStprDn_CnvyrStr AND NOT #sStWtResetRel AND #sSst AND #iqTx_To_Next_0DegTTDown AND NOT #iXferAreaClr_0DegTTDown;
END_REGION

REGION Network 92: STATE Num:250 StWtTTDnStprDn&CnvyrStr
   RUNG wire#powerrail
      Contact( #s250_StWtTTDnStprDn_CnvyrStr )
      wire#w1
      I_Contact( #sStWtResetRel )
      I_Contact( #s250_StWtTTDnStprDn_CnvyrStr_T1 )
      wire#w2
      Coil( #s250_StWtTTDnStprDn_CnvyrStr )
   END_RUNG
   RUNG wire#powerrail
      Contact( #s240_StWtFRTRNxtStnTTDown_T1 )
   END_RUNG wire#w1
   RUNG wire#w2
      { S7_GenerateENO := "TRUE" } Move(in := 250, out1 => #StateNo)
   END_RUNG
   // the same network as SCL:
   #s250_StWtTTDnStprDn_CnvyrStr := (#s250_StWtTTDnStprDn_CnvyrStr OR #s240_StWtFRTRNxtStnTTDown_T1) AND NOT #sStWtResetRel AND NOT #s250_StWtTTDnStprDn_CnvyrStr_T1;
   IF #s250_StWtTTDnStprDn_CnvyrStr THEN #StateNo := 250; END_IF;
END_REGION

REGION Network 93: Actions for STATE Num:250 StWtTTDnStprDn&CnvyrStr
   RUNG wire#powerrail
      Contact( #s250_StWtTTDnStprDn_CnvyrStr )
      wire#w1
      Coil( #qStprDown_TTDown )
   END_RUNG
   RUNG wire#w1
      Coil( #qConvRun_TTDown )
   END_RUNG
   // the same network as SCL:
   #qStprDown_TTDown := #s250_StWtTTDnStprDn_CnvyrStr;
   #qConvRun_TTDown := #s250_StWtTTDnStprDn_CnvyrStr;
END_REGION

REGION Network 94: Transition for STATE Num:260 StWtPalAbsent
   RUNG wire#powerrail
      Contact( #s260_StWtPalAbsent )
      I_Contact( #sStWtResetRel )
      Contact( #sSst )
      I_Contact( #iPalletPrsnt_TTDown )
      Contact( #sPalletAbsntDebTTDown )
      Contact( #iXferAreaClr_0DegTTDown )
      Coil( #s260_StWtPalAbsent_T1 )
   END_RUNG
   // the same network as SCL:
   #s260_StWtPalAbsent_T1 := #s260_StWtPalAbsent AND NOT #sStWtResetRel AND #sSst AND NOT #iPalletPrsnt_TTDown AND #sPalletAbsntDebTTDown AND #iXferAreaClr_0DegTTDown;
END_REGION

REGION Network 95: STATE Num:260 StWtPalAbsent
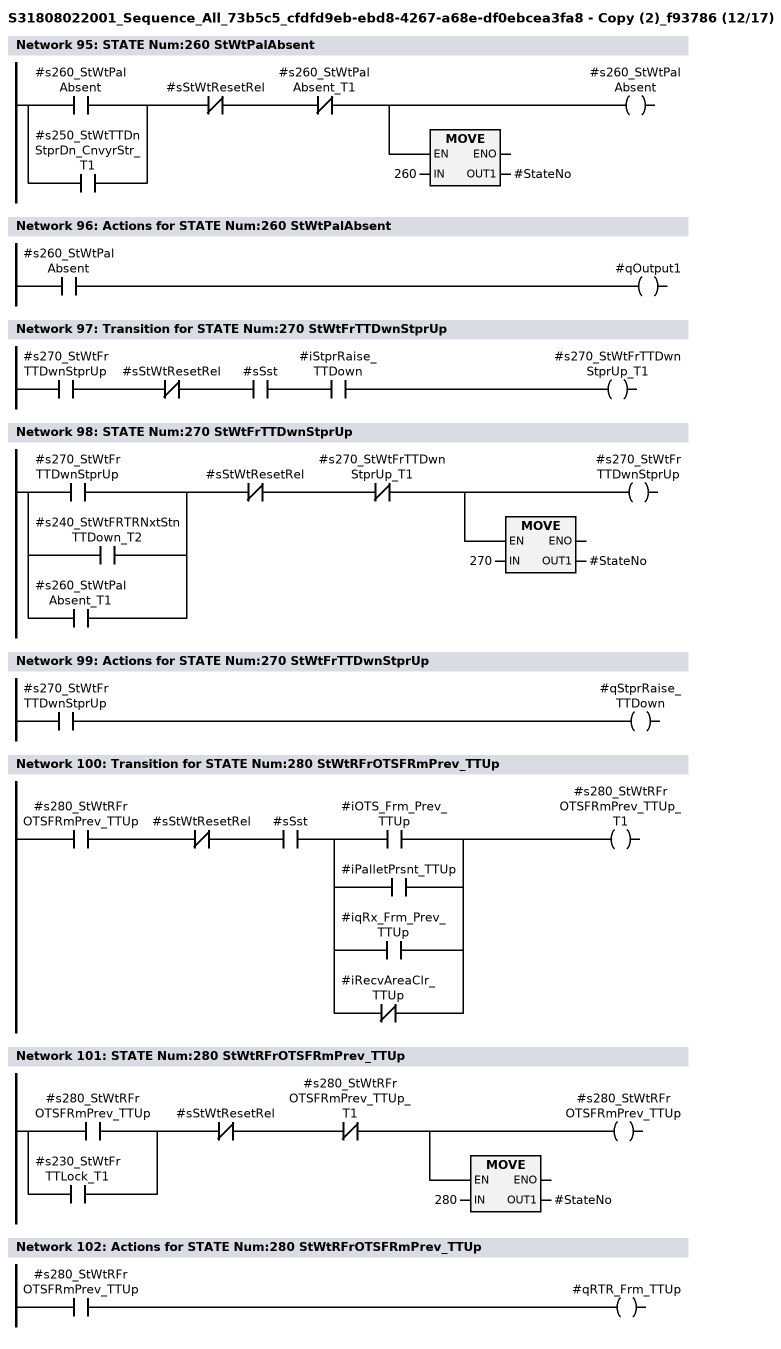
   RUNG wire#powerrail
      Contact( #s260_StWtPalAbsent )
      wire#w1
      I_Contact( #sStWtResetRel )
      I_Contact( #s260_StWtPalAbsent_T1 )
      wire#w2
      Coil( #s260_StWtPalAbsent )
   END_RUNG
   RUNG wire#powerrail
      Contact( #s250_StWtTTDnStprDn_CnvyrStr_T1 )
   END_RUNG wire#w1
   RUNG wire#w2
      { S7_GenerateENO := "TRUE" } Move(in := 260, out1 => #StateNo)
   END_RUNG
   // the same network as SCL:
   #s260_StWtPalAbsent := (#s260_StWtPalAbsent OR #s250_StWtTTDnStprDn_CnvyrStr_T1) AND NOT #sStWtResetRel AND NOT #s260_StWtPalAbsent_T1;
   IF #s260_StWtPalAbsent THEN #StateNo := 260; END_IF;
END_REGION

REGION Network 96: Actions for STATE Num:260 StWtPalAbsent
   RUNG wire#powerrail
      Contact( #s260_StWtPalAbsent )
      Coil( #qOutput1 )
   END_RUNG
   // the same network as SCL:
   #qOutput1 := #s260_StWtPalAbsent;
END_REGION

